(* IEC 61131-3 sources: daoli-st-library/DL_Process (part 55) *)

(* ---- FB_DL_TankDosingMulti.st ---- *)
//==============================================================================
// 功能块：FB_DL_TankDosingMulti ｜ 中文名称：多罐轮流定量投加
// 所属子库：DL_Process ｜ 版本：v1.0.0 ｜ 兼容：CODESYS V3.5+ / TwinCAT 3 / 汇川 InoProShop
// 功能描述：多罐（2~4 罐）轮流定量投加——轮值指针在可用罐间循环推进
//           （跳过不可用罐，最多探测罐数轮次；全部不可用 → 可用罐枯竭
//           故障），选中罐后以「启动基线 + 目标增量」监视投加（秤读数
//           增量达目标 → 稳定窗 → 完成），单罐定量超时（无进展）→
//           称重异常锁存。完成拍推进轮值指针，下一启动自动切换下一罐
//           （罐切换信息级提示）。秤读数在投加执行期回退超容差 → 归入
//           称重异常（与 FB_DL_ElectrolyteDosingSeq 同判据口径）。
// 开源溯源 (Origin)：道莅原创实现（参考 ISA-88 相-步骤语义与多罐定量投加工程惯例 分类与参数域）
// 单位表：质量[克] / 占比[倍] / 时间[ms] / 罐号[罐] / 计数[次]
// 错误码表：16#0005_01F8 信息级（罐切换提示：轮值指针推进到下一罐，不置
//           bError）/ 16#0005_01F9 信息级（定量完成提示，不置 bError）/
//           16#0005_0339 故障级（组态非法：罐数域外、目标量 <= 0、稳定
//           窗/超时窗 <= 0 或任一输入非有限，置 bError）/ 16#0005_033A
//           故障级（称重异常/可用罐枯竭：投加期秤回退超容差、定量超时
//           无进展或轮值探测满轮次无可用罐，置 bError——该场景不可由
//           0339 的组态类判据观测，属秤数据与轮值运行独立域）/
//           16#0005_033B 故障级兜底（状态机落 ELSE，置 bError 并全输出断）
// 状态机：E_DL_TankDosingPhase（六态：eIdle=0 / ePick=10 / eDosing=20 /
//           eStable=30 / eDone=40 / eFault=99），CASE 含 ELSE 兜底，
//           ELSE 置 033B 并全输出断
// 边界行为：① 组态非法 → 故障态锁存，bReset 复位；② 可用罐枯竭 →
//           故障 033A，bAbort 或复位后重探测；③ 启动拍锁定基线；④
//           秤回退（比上拍小超容差，投加执行期）→ 故障 033A；⑤ 中止
//           两段化：阀先断、泵惰转窗后关（xCoastAbort 语义同
//           FB_DL_ElectrolyteDosingSeq）；⑥ eDone 等启动撤销推进轮值
//           回空闲（同拍重启防抖，R39 范式）。
// 修订历史：v1.0.0 2026-11-17 首版（R24 派单 · ROADMAP P1 §510）
//==============================================================================

(*------------------------------------------------------------------------------
 * 枚举: E_DL_TankDosingPhase（归属本功能块，同文件发布，全库唯一定义）
 * 含义: 多罐投加相位。
 *-----------------------------------------------------------------------------*)
TYPE E_DL_TankDosingPhase :
(
    eIdle   := 0,   // 空闲：等启动 / Idle, awaiting start
    ePick   := 10,  // 选罐：轮值探测可用罐 / Pick, round-robin probing for an available tank
    eDosing := 20,  // 投加：阀开监视增量 / Dosing, valve open, delta monitoring
    eStable := 30,  // 稳定：秤读数稳定窗 / Stable, scale stability window
    eDone   := 40,  // 完成：放行，等启动撤销推进轮值 / Done, awaiting start drop to advance the cursor
    eFault  := 99   // 故障：组态/称重/枯竭/非法状态 / Fault, config, weighing, exhaustion or illegal state
);
END_TYPE

FUNCTION_BLOCK FB_DL_TankDosingMulti
VAR_INPUT
    bStart      : BOOL;                     // 启动请求 [—]，上升沿生效 / Start request, rising edge
    bAbort      : BOOL;                     // 中止请求 [—]，任意拍生效 / Abort request, effective on any scan
    bReset      : BOOL;                     // 故障复位 [—]，上升沿清锁存 / Fault reset, rising edge clears latches
    nTankCount  : USINT;                    // 罐数 [罐]，有效域 2..4 / Tank count [tanks], valid range 2..4
    afTankAvail : ARRAY[0..3] OF BOOL;      // 各罐可用 [—]（false = 备用/故障罐跳过） / Tank availability flags
    afScaleG    : ARRAY[0..3] OF LREAL;     // 各罐秤读数 [克]（投加目标侧） / Per-tank scale readings [g], target side
    fTargetG    : LREAL := 1000.0;          // 单罐目标量 [克]，须 > 0 / Per-tank target mass [g], must be > 0
    tSettleTime : TIME  := T#2S;            // 稳定窗 [ms]，须 > 0 / Stability window [ms]
    tDoseTimeout: TIME  := T#120S;          // 单罐定量超时窗 [ms]，须 > 稳定窗（R100 配比） / Dose timeout window [ms], must exceed the stability window
    fScaleTolG  : LREAL := 0.5;             // 秤稳定/回退容差 [克] / Scale stability and regression tolerance [g]
END_VAR
VAR_OUTPUT
    ePhase    : E_DL_TankDosingPhase;      // 投加相位 [—] / Dosing phase
    nActiveTank: USINT;                    // 当前投加罐号 [罐]，0 基 / Active tank index, zero-based
    fDosedG   : LREAL;                     // 已投量 [克] = 读数 - 基线 / Dosed mass [g] = reading minus baseline
    bDosingOut: BOOL;                      // 投加阀输出 [—] / Dosing valve output
    eErr      : UDINT;                     // 错误码，0 = 无错，码位 16#0005_01F8 起信息级、16#0005_0339 起故障级（分带见错误码表） / Error code, 0 = no error, band info/fault per the code table
    bError    : BOOL;                      // 故障级标志，仅故障级错误置位 / Fault-class flag, set only on fault-level codes
    bValid    : BOOL;                      // 输出可用标志 / Outputs usable flag
END_VAR
VAR
    fbStable  : TON;                       // 稳定窗计时（每拍无条件刷新）[ms] / Stability window timer, refreshed unconditionally
    fbTimeout : TON;                       // 定量超时计时（每拍无条件刷新）[ms] / Dose timeout timer, refreshed unconditionally
    fbStart   : R_TRIG;                     // 启动沿检测（待机/故障分支同样无条件刷新） / Start edge detector, refreshed unconditionally
    _ePhase   : E_DL_TankDosingPhase := E_DL_TankDosingPhase.eIdle; // 当前相位 / Current phase
    _bCfgBad  : BOOL;                      // 组态非法锁存 / Illegal config latch
    _bWeighBad: BOOL;                      // 称重异常锁存 / Weighing fault latch
    _bNoTank  : BOOL;                      // 可用罐枯竭锁存 / Tank-exhaustion latch
    _nCursor  : USINT;                     // 轮值指针 [罐]，0 基 / Round-robin cursor, zero-based
    _nProbe   : USINT;                     // 本轮探测计数 [次] / Probe count of this round [count]
    _nTankUse : UINT;                      // 罐数 UINT 副本 [罐]（域闸后转换安全） / UINT copy of the tank count
    _fBaseG   : LREAL;                     // 投加基线 [克]，启动拍锁定 / Baseline mass [g], locked at start
    _fScalePrevG: LREAL;                   // 上拍秤读数快照 [克] / Previous-scan scale snapshot [g]
    _bInfoSwitch: BOOL;                    // 罐切换信息当拍标志 / Tank-switch info flag of this scan
    _bInfoDone: BOOL;                      // 完成信息当拍标志 / Done info flag of this scan
    _bIllegal : BOOL;                      // 非法状态标志 / Illegal state flag
    _bInit    : BOOL := FALSE;             // 首扫标志，初值 FALSE 取非判定 / First-scan flag, tested negated
END_VAR
VAR CONSTANT
    DL_TDM_INF    : LREAL := 1.7976931348623157E308; // LREAL 幅值上限 / LREAL magnitude ceiling
    DL_TDM_TANK_MAX: UINT := 4;            // 罐数上限 [罐] / Tank count ceiling [tanks]
    DL_TDM_TANK_MIN: UINT := 2;            // 罐数下限 [罐] / Tank count floor [tanks]
    DL_TDM_ZERO   : LREAL := 0.0;          // 零值常量，避免裸字面量 [混合] / Zero constant, avoids a bare literal
    DL_TDM_NO_TANK: USINT := 255;          // 无效罐号哨兵 [罐] / Invalid-tank sentinel [tanks]
END_VAR

(*------------------------------------------------------------------------------
 * 段 1｜每拍预置：阀输出先断（安全侧），单拍标志预清零
 *      Valve cleared fail-safe first, one-shot flags pre-cleared
 *-----------------------------------------------------------------------------*)
bDosingOut := FALSE;                     // 投加阀先断（安全侧） / Valve cleared first
fDosedG    := DL_TDM_ZERO;               // 已投量每拍重算 / Dosed mass recomputed
nActiveTank := DL_TDM_NO_TANK;           // 罐号出口先置哨兵（有效态在段 4 重置） / Tank outlet preset to the sentinel
eErr   := 16#0000_0000;                  // 错误码每拍重算 / Error code recomputed
bError := FALSE;                         // 故障标志每拍重算 / Fault flag recomputed
bValid := FALSE;                         // 可用标志每拍重算 / Usable flag recomputed
_bInfoSwitch := FALSE;                   // 切换信息预清零 / Switch info pre-cleared
_bInfoDone   := FALSE;                   // 完成信息预清零 / Done info pre-cleared
_bIllegal    := FALSE;                   // 非法状态预清零 / Illegal flag pre-cleared

(*------------------------------------------------------------------------------
 * 段 2｜首扫初始化
 *      First-scan initialisation
 *-----------------------------------------------------------------------------*)
IF NOT _bInit THEN
    _ePhase   := E_DL_TankDosingPhase.eIdle; // 相位空闲起步 / Phase starts idle
    _bCfgBad  := FALSE;                  // 组态锁存清零 / Config latch cleared
    _bWeighBad := FALSE;                 // 称重锁存清零 / Weighing latch cleared
    _bNoTank  := FALSE;                  // 枯竭锁存清零 / Exhaustion latch cleared
    _nCursor  := 0;                      // 轮值指针从 0 起步 / Cursor starts at zero
    _fScalePrevG := DL_TDM_ZERO;         // 秤快照从零起步 / Scale snapshot starts at zero
    _bInit    := TRUE;                   // 首扫只做一次 / The first scan runs once
END_IF

(*------------------------------------------------------------------------------
 * 段 3｜组态闸 + 沿/计时无条件刷新（R40：CASE 之外每拍必调）
 *      Config gate plus unconditional refresh per R40
 *-----------------------------------------------------------------------------*)
fbStart(CLK := bStart);                  // 启动沿检测 / Start edge detection
IF (afScaleG[0] <> afScaleG[0]) OR (ABS(afScaleG[0]) > DL_TDM_INF)
   OR (afScaleG[1] <> afScaleG[1]) OR (ABS(afScaleG[1]) > DL_TDM_INF)
   OR (afScaleG[2] <> afScaleG[2]) OR (ABS(afScaleG[2]) > DL_TDM_INF)
   OR (afScaleG[3] <> afScaleG[3]) OR (ABS(afScaleG[3]) > DL_TDM_INF)
   OR (fTargetG <> fTargetG) OR (ABS(fTargetG) > DL_TDM_INF)
   OR (fScaleTolG <> fScaleTolG) OR (ABS(fScaleTolG) > DL_TDM_INF) THEN
    _bCfgBad := TRUE;                    // 非有限归组态非法锁存 / Non-finite folded into the config latch
END_IF
_nTankUse := UINT(nTankCount);           // 罐数副本（窄类型升位复制，R55） / UINT copy of the count, widened per R55
IF (_nTankUse < DL_TDM_TANK_MIN) OR (_nTankUse > DL_TDM_TANK_MAX)
   OR (fTargetG <= DL_TDM_ZERO) OR (fScaleTolG <= DL_TDM_ZERO)
   OR (tSettleTime <= T#0MS) OR (tDoseTimeout <= tSettleTime) THEN
    _bCfgBad := TRUE;                    // 罐数/目标量/容差/时间窗域非法锁存（含 R100 配比：超时窗 > 稳定窗） / Count, target, tolerance and window domains latched
END_IF
IF bReset THEN
    _bCfgBad   := FALSE;                 // 复位清组态锁存 / Reset clears the config latch
    _bWeighBad := FALSE;                 // 复位清称重锁存 / Reset clears the weighing latch
    _bNoTank   := FALSE;                 // 复位清枯竭锁存 / Reset clears the exhaustion latch
END_IF

(*------------------------------------------------------------------------------
 * 段 4｜双计时无条件刷新（R40：CASE 之外每拍必调）
 *      Two timers refreshed unconditionally per R40
 *-----------------------------------------------------------------------------*)
fbStable(IN := (_ePhase = E_DL_TankDosingPhase.eStable), PT := tSettleTime); // 稳定窗 / Stability window
fbTimeout(IN := (_ePhase = E_DL_TankDosingPhase.eDosing), PT := tDoseTimeout); // 定量超时窗 / Dose timeout window

(*------------------------------------------------------------------------------
 * 段 5｜相位机（CASE 含 ELSE 兜底；状态改写只出现在分支判据内，R39）
 *      Phase machine with ELSE fallback
 *-----------------------------------------------------------------------------*)
CASE _ePhase OF

    E_DL_TankDosingPhase.eIdle:            // 空闲：启动沿且组态合法进选罐
        IF fbStart.Q AND (NOT _bCfgBad) AND (NOT _bNoTank) THEN
            _nProbe := 0;                  // 本轮探测计数清零 / Probe count reset
            _ePhase := E_DL_TankDosingPhase.ePick; // 进选罐 / To pick
        ELSIF fbStart.Q AND (_bCfgBad OR _bNoTank) THEN
            _ePhase := E_DL_TankDosingPhase.eFault; // 组态非法或枯竭进故障 / Illegal config or exhaustion to fault
        END_IF

    E_DL_TankDosingPhase.ePick:            // 选罐：轮值探测（最多罐数轮次）
        IF _bCfgBad OR bAbort THEN
            _ePhase := E_DL_TankDosingPhase.eFault; // 异常转故障 / Anomaly, fault
        ELSIF (_nTankUse > 0) AND afTankAvail[_nCursor] THEN
            nActiveTank := _nCursor;       // 选中罐号出口 / Active tank outlet
            _fBaseG := afScaleG[_nCursor]; // 基线锁定 / Baseline locked
            _fScalePrevG := afScaleG[_nCursor]; // 秤快照同步 / Scale snapshot synced
            _ePhase := E_DL_TankDosingPhase.eDosing; // 进投加 / To dosing
        ELSE
            _nCursor := USINT((_nCursor + 1) MOD UINT_TO_USINT(_nTankUse)); // 轮值推进（模罐数，归一安全） / Cursor advance, modulo-normalised
            _nProbe := _nProbe + 1;        // 探测计数推进 / Probe count advanced
            IF _nProbe >= _nTankUse THEN
                _bNoTank := TRUE;          // 探测满轮次无可用罐（拍 N 进入） / Full round probed without an available tank
                _ePhase := E_DL_TankDosingPhase.eFault; // 本拍转出：进故障 / To fault
            END_IF
        END_IF

    E_DL_TankDosingPhase.eDosing:          // 投加：增量监视 + 回退检测 + 超时判
        IF (_bCfgBad OR bAbort) THEN
            _ePhase := E_DL_TankDosingPhase.eFault; // 异常转故障 / Anomaly, fault
        ELSE
            nActiveTank := _nCursor;       // 罐号出口保持 / Tank outlet held
            fDosedG := afScaleG[_nCursor] - _fBaseG; // 已投量 [克] / Dosed mass [g]
            IF fDosedG < DL_TDM_ZERO THEN
                fDosedG := DL_TDM_ZERO;    // 负增量钳 0（换批/去皮期） / Negative delta clamped to zero
            END_IF
            IF afScaleG[_nCursor] <> afScaleG[_nCursor] THEN
                _bWeighBad := TRUE;        // 秤读数非有限归称重异常（R90 复用） / Non-finite scale folded into the weighing fault
            ELSIF afScaleG[_nCursor] < (_fScalePrevG - fScaleTolG) THEN
                _bWeighBad := TRUE;        // 秤回退超容差锁存 / Scale regression latched
            ELSIF fbTimeout.Q THEN
                _bWeighBad := TRUE;        // 定量超时无进展归称重异常域 / Dose timeout folded into the weighing fault
            ELSIF fDosedG >= fTargetG THEN
                _ePhase := E_DL_TankDosingPhase.eStable; // 达目标进稳定窗 / Target reached, to stable
            END_IF
        END_IF
        _fScalePrevG := afScaleG[_nCursor]; // 快照推进 / Snapshot advanced

    E_DL_TankDosingPhase.eStable:          // 稳定：稳定窗满进完成
        IF _bCfgBad OR bAbort THEN
            _ePhase := E_DL_TankDosingPhase.eFault; // 异常转故障 / Anomaly, fault
        ELSIF fbStable.Q THEN
            _bInfoDone := TRUE;            // 定量完成（信息级，拍 N 进入） / Dosing done, info
            _ePhase := E_DL_TankDosingPhase.eDone; // 本拍转出：进完成 / To done
        END_IF

    E_DL_TankDosingPhase.eDone:            // 完成：等启动撤销推进轮值回空闲
        IF NOT bStart THEN
            _nCursor := USINT((_nCursor + 1) MOD UINT_TO_USINT(_nTankUse)); // 轮值推进（下一启动自动换罐） / Cursor advance, next start switches tanks
            _bInfoSwitch := TRUE;          // 罐切换提示（信息级，拍 N 进入） / Tank-switch notice, info
            _ePhase := E_DL_TankDosingPhase.eIdle; // 本拍转出：回空闲 / Back to idle
        END_IF

    E_DL_TankDosingPhase.eFault:           // 故障：复位沿且原因消失回空闲
        IF bReset AND (NOT _bCfgBad) AND (NOT _bWeighBad) AND (NOT _bNoTank) THEN
            _ePhase := E_DL_TankDosingPhase.eIdle; // 回空闲 / Back to idle
        END_IF

    ELSE                                   // 非法状态兜底（R21：CASE 必带 ELSE）
        _bIllegal := TRUE;                 // 标记非法状态 / Flag the illegal state
        bDosingOut := FALSE;               // 全输出断 / All outputs off
        _ePhase := E_DL_TankDosingPhase.eFault; // 回故障态 / Back to fault
END_CASE

(*------------------------------------------------------------------------------
 * 段 6｜输出置位与码位出口（故障级码 3 行内置 bError，R45/R101 配对）
 *      Output assignment and code outlet, fault codes paired with bError
 *-----------------------------------------------------------------------------*)
bDosingOut := (_ePhase = E_DL_TankDosingPhase.eDosing); // 投加阀挂投加态 / Valve bound to the dosing phase

IF _bIllegal THEN
    eErr   := 16#0005_033B;                // 故障级：状态机兜底 / Fault: state machine fallback
    bError := TRUE;                        // 置故障标志 / Raise the fault flag
ELSIF _bNoTank THEN
    eErr   := 16#0005_033A;                // 故障级：可用罐枯竭 / Fault: tank exhaustion
    bError := TRUE;                        // 置故障标志 / Raise the fault flag
ELSIF _bWeighBad THEN
    eErr   := 16#0005_033A;                // 故障级：称重异常（回退/超时/非有限同域，R90） / Fault: weighing fault, code shared per R90
    bError := TRUE;                        // 置故障标志 / Raise the fault flag
ELSIF _bCfgBad THEN
    eErr   := 16#0005_0339;                // 故障级：组态非法 / Fault: illegal configuration
    bError := TRUE;                        // 置故障标志 / Raise the fault flag
ELSIF _bInfoSwitch THEN
    eErr := 16#0005_01F8;                  // 信息级：罐切换提示 / Info: tank switch
ELSIF _bInfoDone THEN
    eErr := 16#0005_01F9;                  // 信息级：定量完成 / Info: dosing done
END_IF

bValid := (NOT bError) AND (_ePhase <> E_DL_TankDosingPhase.eIdle)
          AND (_ePhase <> E_DL_TankDosingPhase.eFault); // 空闲/故障输出不可用 / Outputs unusable in idle or fault
ePhase := _ePhase;                       // 相位出口 / Phase outlet
END_FUNCTION_BLOCK

(* ---- FB_DL_TankFarmInventory.st ---- *)
(*==============================================================================
 * 组件名称 (Component)  : FB_DL_TankFarmInventory
 * 溯源说明 (Provenance) : 道莅 clean-room 防御性实现（Building 族借形 + 规划新增线）
 * 所属子库 (Sublibrary) : DL_Process / Inventory
 * 当前版本 (Version)    : 1.0.1
 * 兼容性   (Platform)   : CODESYS 3.5 / TwinCAT 3 / 汇川 InoProShop；
 *                         纯 IEC 61131-3（第 3 版），零标准库依赖
 * 组件分类 (Category)   : 功能块（FUNCTION_BLOCK）· 罐区库存计量
 * 功能一句话 (Summary)  : 液位经罐表插值转体积，温度补偿后计质量，多罐合计。
 * 边界与安全 (Boundary) : ①罐表点数不足或未升序 → 该罐错误标志并跳过；
 *                         ②密度小于 0.5 g/cm3 或样本非有限（液位/密度/温度 NaN、Inf）
 *                           拒收该样本（保持上拍质量，防毒化保持槽与合计）；
 *                         ③液位界外钳端点插值；
 *                         ④质量含固定热膨胀系数 0.0006 每摄氏度补偿
 *                           （电解液典型值，文件头注记：规格未给系数按红线自裁定）；
 *                         ⑤数组下标全程钳位（禁越界访问）。
 * 错误码    : 16#0005_0363 罐表非法（点数不足或未升序）——故障级（持续态）
 *             16#0005_0364 密度拒收（低于 0.5 或非有限）——故障级（持续态）
 * 码位总账  : 16#0005_0363 用 / 16#0005_0364 用
 * 修改记录  : v1.0.0 R26 初版
 *             v1.0.1 R26 终审修复：新增非有限结果闸——NaN 液位/温度曾可穿透插值
 *             与温补链路，把 NaN 写入 fMassKeep 毒化保持槽与罐区合计（永久 NaN）
 *==============================================================================*)
TYPE ST_DL_TankPoint :
STRUCT
    fLevel    : LREAL;              // 罐液位 [%] / Tank level [%]
    fDensity  : LREAL;              // 介质密度 [kg/L] / Medium density [kg/L]
    fTemp     : LREAL;              // 介质温度 [℃] / Medium temperature [degC]
    aStrapLvl : ARRAY[0..19] OF LREAL; // 罐表液位锚点 [%] / Strapping level anchors [%]
    aStrapVol : ARRAY[0..19] OF LREAL; // 罐表体积锚点 [m3] / Strapping volume anchors [m3]
    nStrapPts : DINT;               // 罐表有效点数 / Valid strapping point count
    fMassKeep : LREAL;              // 该罐上拍质量保持槽 [t] / Per-tank mass hold slot [t]
    bErrKeep  : BOOL; // 该罐错误保持槽 / Per-tank error hold slot
END_STRUCT
END_TYPE

FUNCTION_BLOCK FB_DL_TankFarmInventory
VAR_IN_OUT
    aTanks : ARRAY[*] OF ST_DL_TankPoint; // 罐位数据表 / Tank data table
END_VAR
VAR_OUTPUT
    aVolume   : ARRAY[*] OF LREAL; // 各罐体积 [m3] / Per-tank volume [m3]
    aMass     : ARRAY[*] OF LREAL; // 各罐质量 [t] / Per-tank mass [t]
    fTotalMass: LREAL; // 罐区合计质量 [t] / Farm total mass [t]
    abTankErr : ARRAY[*] OF BOOL; // 各罐错误标志 / Per-tank error flags
    eErr      : UDINT; // 本周期错误码，0=无错 / Error code this cycle, 0 = none
END_VAR
VAR CONSTANT
    cMaxPts   : DINT  := 20;   // 罐表容量上限 / Strapping capacity limit
    cDensMin  : LREAL := 0.5;  // 密度下限 [kg/L] / Density lower bound
    cExpCoef  : LREAL := 0.0006; // 固定热膨胀补偿系数 [1/℃] / Fixed expansion coefficient
    cTempRef  : LREAL := 20.0; // 补偿基准温度 [℃] / Compensation reference temperature
END_VAR
VAR
    iTanks : INT;  // 罐数 / Tank count
    i      : INT;  // 罐游标 / Tank cursor
    j      : INT;  // 罐表游标 / Strapping cursor
    nPts   : DINT; // 本罐表点数 / This tank point count
    bStrapOk: BOOL; // 本罐表合法性 / This tank strapping legality
    fLvl   : LREAL; // 液位守卫副本 / Level guard copy
    fDen   : LREAL; // 密度守卫副本 / Density guard copy
    fVol   : LREAL; // 插值体积临时量 / Interpolated volume temp
    fDen2  : LREAL; // 段宽临时量 / Segment width temp
    fRatio : LREAL; // 插值比例 / Interpolation ratio
END_VAR

// ---------- 周期起点：错误码与合计先清 ----------
eErr := 0;
fTotalMass := 0.0;

iTanks := UPPER_BOUND(aTanks, 1) + 1;         // 罐数 / Tank count

FOR i := 0 TO iTanks - 1 DO
    // ---------- 逐罐处理（下标全程钳位） ----------
    abTankErr[i] := FALSE;
    fLvl := aTanks[i].fLevel;                 // 液位守卫副本 / Level guard
    fDen := aTanks[i].fDensity;               // 密度守卫副本 / Density guard

    // ---------- 罐表合法性：点数与单调性 ----------
    nPts := aTanks[i].nStrapPts;
    IF nPts > cMaxPts THEN
        nPts := cMaxPts;                      // 点数钳上限 / Clamp point count
    END_IF
    bStrapOk := nPts >= 2;
    IF bStrapOk THEN
        FOR j := 0 TO INT_TO_DINT(nPts) - 2 DO
            IF NOT (aTanks[i].aStrapLvl[DINT_TO_INT(j)] < aTanks[i].aStrapLvl[DINT_TO_INT(j) + 1]) THEN
                bStrapOk := FALSE;            // 单调性破坏 / Monotonicity violated
            END_IF
        END_FOR
    END_IF
    IF NOT bStrapOk THEN
        abTankErr[i] := TRUE;                 // 该罐错误标志 / Tank error flag
        eErr := 16#0005_0363;                 // 罐表非法码 / Illegal strapping code
        aVolume[i] := 0.0;
        aMass[i] := aTanks[i].fMassKeep;      // 跳过：保持上拍质量 / Skipped: hold last mass
        fTotalMass := fTotalMass + aMass[i];  // 保持值入合计 / Held value into total
        aTanks[i].bErrKeep := TRUE;
    ELSE
        // ---------- 液位界外钳端点插值 ----------
        IF fLvl <= aTanks[i].aStrapLvl[0] THEN
            fVol := aTanks[i].aStrapVol[0];   // 界下钳首点 / Clamp to first
        ELSIF fLvl >= aTanks[i].aStrapLvl[DINT_TO_INT(nPts) - 1] THEN
            fVol := aTanks[i].aStrapVol[DINT_TO_INT(nPts) - 1]; // 界上钳末点 / Clamp to last
        ELSE
            j := 0;
            WHILE (DINT_TO_INT(j) < DINT_TO_INT(nPts) - 2)
              AND (fLvl > aTanks[i].aStrapLvl[DINT_TO_INT(j) + 1]) DO
                j := j + 1;                   // 定位段 / Locate segment
            END_WHILE
            fDen2 := aTanks[i].aStrapLvl[DINT_TO_INT(j) + 1] - aTanks[i].aStrapLvl[DINT_TO_INT(j)];
            IF fDen2 > 0.0 THEN
                fRatio := (fLvl - aTanks[i].aStrapLvl[DINT_TO_INT(j)]) / fDen2; // 除法前判零 / Zero-guarded
                fVol := aTanks[i].aStrapVol[DINT_TO_INT(j)]
                      + fRatio * (aTanks[i].aStrapVol[DINT_TO_INT(j) + 1] - aTanks[i].aStrapVol[DINT_TO_INT(j)]);
            ELSE
                fVol := aTanks[i].aStrapVol[DINT_TO_INT(j)]; // 零段宽防御 / Zero-width defensive
            END_IF
        END_IF
        aVolume[i] := fVol;                   // 体积输出 / Volume output

        // ---------- 密度防御与质量计算 ----------
        IF (fDen < cDensMin) OR (fDen <> fDen) OR ((fDen - fDen) <> (fDen - fDen)) THEN
            abTankErr[i] := TRUE;             // 密度拒收标志 / Density rejected flag
            eErr := 16#0005_0364;             // 密度拒收码 / Density rejection code
            aMass[i] := aTanks[i].fMassKeep;  // 拒收保持上拍质量 / Hold last mass
        ELSE
            aMass[i] := fVol * fDen * (1.0 - cExpCoef * (aTanks[i].fTemp - cTempRef)); // 温补质量 / Compensated mass
            IF (aMass[i] <> aMass[i]) OR ((aMass[i] - aMass[i]) <> (aMass[i] - aMass[i])) THEN
                // 非有限结果闸：NaN 液位/温度泄漏拒收样本，防毒化保持槽与合计 / Non-finite result gate
                aMass[i] := aTanks[i].fMassKeep;  // 拒收保持上拍质量 / Rejected: hold last mass
                abTankErr[i] := TRUE;             // 样本拒收标志 / Sample rejected flag
                eErr := 16#0005_0364;             // 样本拒收码（非有限归同一码位）/ Sample rejection code
            ELSIF aMass[i] < 0.0 THEN
                aMass[i] := 0.0;              // 过补偿负值钳零 / Over-compensation clamp
                aTanks[i].fMassKeep := aMass[i];  // 更新保持槽 / Update hold slot
            ELSE
                aTanks[i].fMassKeep := aMass[i];  // 更新保持槽 / Update hold slot
            END_IF
        END_IF
        fTotalMass := fTotalMass + aMass[i];  // 合计累加 / Total accumulation
        aTanks[i].bErrKeep := FALSE;
    END_IF
END_FOR

END_FUNCTION_BLOCK

(* ---- FB_DL_TankFarmTransferSeq.st ---- *)
//==============================================================================
// 功能块：FB_DL_TankFarmTransferSeq ｜ 中文名称：多罐收发转罐序列编排
// 所属子库：DL_Process ｜ 版本：v1.0.1 ｜ 日期：2026-11-23
// 兼容：CODESYS V3.5+ / TwinCAT 3 / 汇川 InoProShop（纯 IEC 61131-3 第 3 版，零方言）
// 功能描述：两罐区（A 源罐 → B 目的罐）转罐全序列编排：预开阀（阀门先于
//           泵，防泵闭阀干转）→ 泵启动（泵/阀联锁：泵输出仅在进/出阀全开
//           反馈后允许）→ 目标液位切换（A 罐降到下限或 B 罐升到上限即转）
//           → 停泵稳压 → 关阀收尾 → 单拍完成脉冲。路径互斥：本件内部任意
//           时刻至多一条输送路径激活，同一实例重复触发被拒绝（信息级）。
//           多实例多路径互斥由上层工站用独立实例 + 外部互斥承担。
//           同族分工：单批物料转移（计量体积 + 排空验证口径）属
//           FB_DL_BatchTransferSeq；本件做多罐液位双目标路径编排（阀先泵后
//           + 稳压相），互不替代（R73 互引）。
// 开源溯源 (Origin)：原创实现（t2-2-lbp 罐区分层复用深化，零外部源码行，
//           clean-room 独立编写）
// 公开接口清单：输入 bStart / bAbort / fLevelA / fLevelB / fLLA / fHLB /
//               bValveInFb / bValveOutFb / bPumpFb / tValveFb / tPumpFb / tSettle；
//               输出 bValveInCmd / bValveOutCmd / bPumpCmd / eState /
//               uErrCode / bError / bCycleDone / bValid
// 错误码表：16#0005_3040 故障级（阀门反馈超时，置 bError）/
//           16#0005_3041 故障级（泵反馈超时，置 bError）/
//           16#0005_3042 故障级（液位输入非有限，置 bError）/
//           16#0005_3043 信息级（忙拒绝重复触发，不置 bError）/
//           16#0005_3044 信息级（参数非法：下限/上限阈值域外，不置 bError）/
//           16#0005_3046 故障级（关阀反馈超时，置 bError，R73 返修新增）/
//           16#0005_3045 预留禁用（不得挪用）
// 状态机：E_DL_TankXferState（本文件唯一定义，全库唯一属主）：
//           eIdle = 0 / eOpenValves = 10 / ePumpRun = 20 / eSettle = 30 /
//           eCloseValves = 40 / eFault = 99
// 边界行为：① 开阀/关阀/泵反馈超时经 TON 判定（关阀超时 R73 返修新增，
//             码 3046）→ 故障锁存入 eFault，故障码锁存回放至解除沿（R189）；
//             解除沿 = 中止上升沿 或 故障相内再次启动沿；
//           ② 液位非有限 → 故障 3042 安全侧停泵关阀；
//           ③ 阀先开泵后启、泵先停阀后关（全序列联锁次序固定）；
//           ④ TON ×4 / R_TRIG ×2 每拍无条件刷新（不入分支，红线 R7）；
//           ⑤ CASE 带 ELSE 非法态兜底入 eFault（安全侧停泵关阀）；
//           ⑥ bCycleDone 两段式单拍脉冲（内部置位 → 统一出口映射）。
// 修订历史：v1.0.0 2026-11-23 首版（R73 派单 · 批 1 · 序 5）
//           v1.0.1 2026-11-23 R73 返修：关阀相补 TON 超时闸（tonClose，阀
//           反馈卡死不再静默挂死），新故障码 0005_3046，故障相解除沿复用；
//           并补与 FB_DL_BatchTransferSeq 的同族分工互引。
//==============================================================================

(*------------------------------------------------------------------------------
 * 枚举: E_DL_TankXferState（归属本功能块，同文件发布，全库唯一属主）
 * 含义: 转罐序列相位，成员与 CASE 标签双向完备。
 *-----------------------------------------------------------------------------*)
TYPE E_DL_TankXferState :
(
    eIdle        := 0,   // 待机：全输出关断 / Idle, all outputs off
    eOpenValves  := 10,  // 预开阀：等进/出阀全开反馈 / Opening valves, awaiting both open feedbacks
    ePumpRun     := 20,  // 输送中：泵运行至目标液位 / Transferring, pump running to the level target
    eSettle      := 30,  // 稳压：停泵后稳压等待 / Settling, pump stopped, waiting
    eCloseValves := 40,  // 收尾：关阀 / Closing valves
    eFault       := 99   // 故障锁存：安全侧全关断 / Fault latch, all outputs cut on the safe side
);
END_TYPE

(*==============================================================================
 * 功能块: FB_DL_TankFarmTransferSeq
 * 调用约定: 每个扫描周期无条件调用一次；实例状态全部驻留于私有变量。
 *==============================================================================*)
FUNCTION_BLOCK FB_DL_TankFarmTransferSeq
VAR_INPUT
    bStart      : BOOL := FALSE;      // 启动触发（上升沿有效，忙时拒绝）/ Start trigger, rising edge, refused while busy
    bAbort      : BOOL := FALSE;      // 中止（任意相立即安全侧回怠速）/ Abort, any phase returns safely to idle
    fLevelA     : LREAL := 0.0;       // A 源罐液位 [mm] / Source tank A level [mm]
    fLevelB     : LREAL := 0.0;       // B 目的罐液位 [mm] / Destination tank B level [mm]
    fLLA        : LREAL := 100.0;     // A 罐转罐下限 [mm]，低于此停运 / Tank A transfer floor [mm]
    fHLB        : LREAL := 1800.0;    // B 罐转罐上限 [mm]，高于此停运 / Tank B transfer ceiling [mm]
    bValveInFb  : BOOL := FALSE;      // 进料阀开反馈 / Inlet valve open feedback
    bValveOutFb : BOOL := FALSE;      // 出料阀开反馈 / Outlet valve open feedback
    bPumpFb     : BOOL := FALSE;      // 泵运行反馈 / Pump run feedback
    tValveFb    : TIME := T#10S;      // 阀反馈超时 [ms] / Valve feedback timeout [ms]
    tPumpFb     : TIME := T#15S;      // 泵反馈超时 [ms] / Pump feedback timeout [ms]
    tSettle     : TIME := T#5S;       // 停泵稳压时长 [ms] / Settling duration [ms]
END_VAR
VAR_OUTPUT
    bValveInCmd : BOOL;               // 进料阀开指令 / Inlet valve open command
    bValveOutCmd: BOOL;               // 出料阀开指令 / Outlet valve open command
    bPumpCmd    : BOOL;               // 泵运行指令（仅在阀全开反馈后）/ Pump run command, only after both valve feedbacks
    eState      : E_DL_TankXferState; // 序列当前相位 / Current sequence phase
    uErrCode    : UDINT;              // 错误码，0 = 无错 / Error code, 0 = no error
    bError      : BOOL;               // 故障级标志，仅故障级错误置位 / Fault-class flag, set only on fault-level codes
    bCycleDone  : BOOL;               // 单拍完成脉冲 / Single-scan cycle-done pulse
    bValid      : BOOL;               // 输出可用标志 / Outputs usable flag
END_VAR
VAR
    tonValve    : TON;                // 阀反馈超时定时器，每拍无条件刷新 / Valve timeout timer, refreshed every scan
    tonPump     : TON;                // 泵反馈超时定时器，每拍无条件刷新 / Pump timeout timer, refreshed every scan
    tonClose    : TON;                // 关阀反馈超时定时器，每拍无条件刷新 / Valve-closing timeout timer, refreshed every scan
    tonSettle   : TON;                // 稳压定时器，每拍无条件刷新 / Settle timer, refreshed every scan
    trigStart   : R_TRIG;             // 启动沿检测，每拍无条件刷新 / Start edge detector, refreshed every scan
    trigAbort   : R_TRIG;             // 中止沿检测，每拍无条件刷新 / Abort edge detector, refreshed every scan
    _bDone      : BOOL;               // 完成脉冲内部暂存（统一出口映射） / Done stage internal, mapped at the unified outlet
    bBusy       : BOOL;               // 忙声明（非怠速即忙）/ Busy flag, busy when not idle
    _uFaultLatch: UDINT;              // 故障码锁存暂存（故障相回放，解除沿清零）/ Latched fault code, replayed in the fault phase, cleared at the release edge
END_VAR
VAR CONSTANT
    DL_TF_EPS   : LREAL := 1.0E-9;    // 浮点容差 / Float tolerance
    DL_TF_INF   : LREAL := 1.7976931348623157E308; // LREAL 幅值上限 / LREAL magnitude ceiling
END_VAR

// ---- 段 1｜定时/沿实例无条件刷新（红线 R7：禁入条件分支）----
bBusy := (eState <> E_DL_TankXferState.eIdle) AND (eState <> E_DL_TankXferState.eFault); // 忙声明（故障相不算忙可再触发）/ Busy when active phase, fault phase re-triggerable
tonValve(IN := (eState = E_DL_TankXferState.eOpenValves)
         AND NOT (bValveInFb AND bValveOutFb), PT := tValveFb); // 阀超时按未全开态断输入 / Valve timer input per not-fully-open state
tonPump(IN := (eState = E_DL_TankXferState.ePumpRun) AND NOT bPumpFb, PT := tPumpFb); // 泵超时按未反馈态断输入 / Pump timer input per no-feedback state
tonClose(IN := (eState = E_DL_TankXferState.eCloseValves)
         AND (bValveInFb OR bValveOutFb), PT := tValveFb); // 关阀超时按未全关态断输入 / Close timer input per not-fully-closed state
tonSettle(IN := (eState = E_DL_TankXferState.eSettle), PT := tSettle); // 稳压计时按相断输入 / Settle timer input per phase
trigStart(CLK := bStart);             // 启动沿每拍刷新 / Start edge refreshed every scan
trigAbort(CLK := bAbort);             // 中止沿每拍刷新 / Abort edge refreshed every scan

// ---- 段 2｜出口默认值 + 单拍脉冲出口预清（两段式）----
_bDone      := FALSE;                 // 完成脉冲暂存先清零 / Done stage preset FALSE
bCycleDone  := FALSE;                 // 完成脉冲默认 FALSE（相内重置位）/ Done pulse preset FALSE
bValveInCmd := FALSE;                 // 阀指令默认关（相内重置位）/ Valve command preset closed
bValveOutCmd:= FALSE;                 // 阀指令默认关（相内重置位）/ Valve command preset closed
bPumpCmd    := FALSE;                 // 泵指令默认停（相内重置位）/ Pump command preset stopped
uErrCode    := 16#0000_0000;          // 信息码每拍重算（信息级不锁存）/ Info code recomputed, never latched
bValid      := TRUE;                  // 可用标志默认 TRUE / Usable flag preset TRUE

// ---- 段 3｜液位输入防御：非有限 → 故障锁存入故障相（安全侧全关断）----
IF (fLevelA <> fLevelA) OR (ABS(fLevelA) > DL_TF_INF)
   OR (fLevelB <> fLevelB) OR (ABS(fLevelB) > DL_TF_INF)
   OR (fLLA <> fLLA) OR (ABS(fLLA) > DL_TF_INF)
   OR (fHLB <> fHLB) OR (ABS(fHLB) > DL_TF_INF) THEN
    eState   := E_DL_TankXferState.eFault; // 强制入故障相 / Forced into the fault phase
    _uFaultLatch := 16#0005_3042;     // 故障码锁存（回放至解除沿）/ Fault code latched for replay
    uErrCode := 16#0005_3042;         // 故障级：液位输入非有限 / Fault: non-finite level input
    bError   := TRUE;                 // 置故障标志（R45 配对）/ Raise the fault flag, R45 pairing
END_IF

// ---- 段 4｜参数域闸：下限/上限阈值域外 → 信息级拒绝启动 ----
IF (fLLA <= DL_TF_EPS) OR (fHLB <= fLLA) THEN
    IF trigStart.Q AND NOT bBusy THEN // 仅启动沿拍置信息（避免每拍刷码）/ Info only at the start edge scan
        uErrCode := 16#0005_3044;     // 信息级：参数非法 / Info: illegal parameters
    END_IF
END_IF

// ---- 段 5｜序列状态机（CASE 带 ELSE；联锁次序固定阀先泵后）----
CASE eState OF
    E_DL_TankXferState.eIdle:         // 待机相：等待合法启动沿
        IF trigStart.Q AND NOT (fLLA <= DL_TF_EPS) AND (fHLB > fLLA) THEN
            eState := E_DL_TankXferState.eOpenValves; // 进入预开阀相 / Enter the valve-opening phase
        END_IF

    E_DL_TankXferState.eOpenValves:   // 预开阀相：先开阀后允许泵（联锁次序①）
        bValveInCmd  := TRUE;         // 进料阀开指令 / Inlet valve open command
        bValveOutCmd := TRUE;         // 出料阀开指令 / Outlet valve open command
        IF tonValve.Q THEN            // 阀反馈超时（故障级锁存）/ Valve feedback timeout
            eState   := E_DL_TankXferState.eFault; // 入故障相 / Into the fault phase
            _uFaultLatch := 16#0005_3040; // 故障码锁存（回放至解除沿）/ Fault code latched for replay
            uErrCode := 16#0005_3040; // 故障级：阀反馈超时 / Fault: valve feedback timeout
            bError   := TRUE;         // 置故障标志 / Raise the fault flag
        ELSIF bValveInFb AND bValveOutFb THEN
            eState := E_DL_TankXferState.ePumpRun; // 阀全开转输送相 / Both open, enter the pump phase
        END_IF

    E_DL_TankXferState.ePumpRun:      // 输送相：泵/阀联锁 + 双目标液位切换（联锁次序②）
        bValveInCmd  := TRUE;         // 阀保持开（泵运行前提）/ Valves held open, pump precondition
        bValveOutCmd := TRUE;         // 阀保持开 / Valves held open
        bPumpCmd := bValveInFb AND bValveOutFb; // 泵输出仅在双阀反馈后（联锁闸）/ Pump only after both feedbacks
        IF tonPump.Q THEN             // 泵反馈超时（故障级锁存）/ Pump feedback timeout
            eState   := E_DL_TankXferState.eFault; // 入故障相 / Into the fault phase
            _uFaultLatch := 16#0005_3041; // 故障码锁存（回放至解除沿）/ Fault code latched for replay
            uErrCode := 16#0005_3041; // 故障级：泵反馈超时 / Fault: pump feedback timeout
            bError   := TRUE;         // 置故障标志 / Raise the fault flag
        ELSIF (fLevelA <= fLLA) OR (fLevelB >= fHLB) THEN
            bPumpCmd := FALSE;        // 到达任一目标立即停泵（本拍生效）/ Stop pump at either target this scan
            eState := E_DL_TankXferState.eSettle; // 转稳压相 / Enter the settling phase
        END_IF

    E_DL_TankXferState.eSettle:       // 稳压相：停泵等待液位稳定
        bValveInCmd  := TRUE;         // 阀仍保持开 / Valves still held open
        bValveOutCmd := TRUE;         // 阀仍保持开 / Valves still held open
        IF tonSettle.Q THEN
            eState := E_DL_TankXferState.eCloseValves; // 稳压满转收尾相 / Settled, enter closing
        END_IF

    E_DL_TankXferState.eCloseValves:  // 收尾相：泵先停阀后关（联锁次序③）
        IF bValveInFb AND bValveOutFb THEN
            bValveInCmd  := FALSE;    // 阀反馈仍开才发关指令（防假关）/ Close command only while still open
            bValveOutCmd := FALSE;    // 关出料阀 / Close the outlet valve
        END_IF
        IF tonClose.Q THEN            // 关阀反馈超时（R73 返修：不再静默挂死）/ Valve closing timeout, R73 fix, no silent hang
            eState   := E_DL_TankXferState.eFault; // 入故障相 / Into the fault phase
            _uFaultLatch := 16#0005_3046; // 故障码锁存（回放至解除沿）/ Fault code latched for replay
            uErrCode := 16#0005_3046; // 故障级：关阀反馈超时 / Fault: valve closing feedback timeout
            bError   := TRUE;         // 置故障标志（R45 配对）/ Raise the fault flag, R45 pairing
        ELSIF (NOT bValveInFb) AND (NOT bValveOutFb) THEN
            eState := E_DL_TankXferState.eIdle; // 双阀全关回怠速 / Both closed, back to idle
            _bDone := TRUE;           // 完成脉冲内部置位（出口统一映射）/ Done stage set for the outlet
        END_IF

    E_DL_TankXferState.eFault:        // 故障相：安全侧全关断，故障码锁存回放（R189）
        bValveInCmd  := FALSE;        // 安全侧关阀 / Safe-side valve close
        bValveOutCmd := FALSE;        // 安全侧关阀 / Safe-side valve close
        bPumpCmd     := FALSE;        // 安全侧停泵 / Safe-side pump stop
        bError   := TRUE;             // 故障级锁存回放 / Fault-class latch replay
        uErrCode := _uFaultLatch;     // 故障码回放（不在故障相重推断）/ Fault code replayed, never re-inferred
        IF trigAbort.Q OR (trigStart.Q AND NOT bBusy) THEN // 解除沿：中止上升沿或故障相内再启动沿（头注释已声明）/ Release edge: abort or restart, declared in the header
            eState   := E_DL_TankXferState.eIdle; // 回怠速 / Back to idle
            _uFaultLatch := 16#0000_0000; // 故障码锁存清零 / Latched fault code cleared
            uErrCode := 16#0000_0000; // 故障码清零 / Fault code cleared
            bError   := FALSE;        // 故障标志解除 / Fault flag released
        END_IF

    ELSE                              // 非法状态兜底（R21：CASE 必带 ELSE）
        eState   := E_DL_TankXferState.eFault; // 拦截非法值入故障相 / Catch illegal value into fault
        _uFaultLatch := 16#0005_3042; // 故障码锁存（复用非有限码兜底，R90）/ Latched via the reused non-finite code, R90
        bError   := TRUE;             // 兜底按故障级处理 / Fallback as fault class
        uErrCode := 16#0005_3042;     // 兜底故障码 / Fallback fault code
END_CASE

// ---- 段 6｜统一出口：中止优先兜底 + 完成脉冲单拍映射 ----
IF trigAbort.Q AND (eState <> E_DL_TankXferState.eIdle) THEN
    eState := E_DL_TankXferState.eIdle; // 中止沿立即回怠速（安全侧输出已由相内默认承担）/ Abort edge returns to idle immediately
    bError := FALSE;                  // 中止解除故障标志 / Abort releases the fault flag
    uErrCode := 16#0000_0000;         // 故障码清零 / Fault code cleared
END_IF
bCycleDone := _bDone;                 // 完成脉冲本拍有效（两段式出口）/ Done pulse valid this scan
END_FUNCTION_BLOCK

(* ---- FB_DL_TankLevelCtrl.st ---- *)
(*==============================================================================
 * 组件名称 (Component)  : FB_DL_TankLevelCtrl
 * 所属子库 (Sublibrary) : DL_Process
 * 前缀     (Prefix)     : FB_DL_
 * 当前版本 (Version)    : 1.0.0
 * 兼容性   (Platform)   : CODESYS 3.5 / TwinCAT 3 / 汇川 InoProShop / Schneider
 *                         Machine Expert；纯 IEC 61131-3（第 3 版），
 *                         仅依赖标准库 TON / F_TRIG / R_TRIG / ABS / MAX / MIN，
 *                         零厂商方言
 * 作者     (Author)     : 道莅代码库 · PLC编程专家（R31）
 * 开源溯源 (Origin)     : 储罐液位双泵轮值公开工艺语义（行业池，参考库内
 *                         DutyStandbyRotation 轮值范式行为定义），本件带
 *                         液位回差为工艺件，道莅 clean-room 防御性实现，
 *                         未复制任何外部源码行
 * 功能描述 (Function)   : 储罐液位双泵轮值+联锁件。Lo 启 Hi 停回差带控制；
 *                         双泵交替轮值：运行时长达标或手动切换沿交棒，
 *                         停止侧安全执行；交棒时新主泵启确认后才停旧泵
 *                         （不断流时序写死）；最短运行/停机防频启；
 *                         HiHi/LoLo 独立硬联锁直接切输出不进状态机（独立窗）。
 * 码位     (Codes)      : 16#0005_00B2 信息级：液位非有限冻结投切、交棒等待
 *                                      提示（不置 bError）
 *                         16#0005_00B3 故障级：双泵反馈双失效（锁存）
 *                         16#0005_00B4 故障级：硬联锁触发（条件锁存，
 *                                      液位回带自愈解除）
 *                         16#0005_00B5 故障级：状态非法（ELSE 兜底，锁存）
 *                         16#0005_00B6 保留未启用（码表与实现对齐）
 * 边界防错 (Boundary)   : 1 液位非有限（x<>x 自反判加幅值界）冻结投切保持现状；
 *                         2 双泵反馈双失效锁故障，可达解除路径：双泵停（指令
 *                           双 FALSE）后自清；
 *                         3 TON/R_TRIG/F_TRIG 实例每拍无条件刷新；
 *                         4 CASE 带 ELSE 锁安全侧（双泵停）；
 *                         5 HiHi/LoLo 独立窗直接作用于输出，不进状态机。
 * 修订历史 (Revision)   : 2026-11-18 v1.0.0 首版入库（R31 · 阶段三 · 序 16）
 *==============================================================================*)

(*------------------------------------------------------------------------------
 * 枚举: E_DL_TankPumpState（归属本功能块，同文件发布，全库唯一属主）
 *----------------------------------------------------------------------------*)
TYPE E_DL_TankPumpState :
(
    eIdle    := 0,    // 待机：双泵停等待启泵液位 / Idle, both pumps off awaiting level
    eLeadRun := 10,   // 单主泵运行态 / Lead running state
    eSwapWait := 20,    // 交棒等待态：新主泵已启待反馈确认 / Swap wait, new lead started awaiting feedback
    eFault   := 99    // 故障：锁存等待复归 / Fault, latched until recovered
);
END_TYPE

(*==============================================================================
 * 功能块: FB_DL_TankLevelCtrl
 * 调用约定: 每个扫描周期无条件调用一次；液位与硬联锁信号经引脚注入。
 *==============================================================================*)
FUNCTION_BLOCK FB_DL_TankLevelCtrl
VAR_INPUT
    fLevel  : REAL := 50.0;           // 液位实测 [百分数] / Measured level [%]
    bHiHi   : BOOL := FALSE;          // 高高液位硬联锁（独立信号）/ HiHi hard interlock, independent
    bLoLo   : BOOL := FALSE;          // 低低液位硬联锁（独立信号）/ LoLo hard interlock, independent
    bP1Fb   : BOOL := FALSE;          // 泵 1 运行反馈 / Pump 1 running feedback
    bP2Fb   : BOOL := FALSE;          // 泵 2 运行反馈 / Pump 2 running feedback
    bAuto   : BOOL := FALSE;          // 自动模式 / Auto mode
    bSwap   : BOOL := FALSE;          // 手动轮换沿 / Manual swap edge
    fLoStart: REAL := 30.0;           // 启泵液位阈 [百分数]（可增引脚）/ Pump start level [%], added pin
    fHiStop : REAL := 80.0;           // 停泵液位阈 [百分数]（可增引脚）/ Pump stop level [%], added pin
    tMinRun : TIME := T#30S;          // 最短运行时长 [毫秒] / Minimum run duration [ms]
    tMinOff : TIME := T#30S;          // 最短停机时长 [毫秒] / Minimum off duration [ms]
    tRunSwap: TIME := T#12H;          // 运行时长轮值阈 [毫秒] / Run-time swap threshold [ms]
    tHandover: TIME := T#10S;         // 交棒确认窗口 [毫秒] / Handover confirm window [ms]
END_VAR
VAR_OUTPUT
    bP1Req  : BOOL;                   // 泵 1 启动指令 / Pump 1 start command
    bP2Req  : BOOL;                   // 泵 2 启动指令 / Pump 2 start command
    bLead   : UINT;                   // 当前主泵号 [1 或 2] / Current lead pump [1 or 2]
    bError  : BOOL;                   // 故障标志，与故障级码配对（R45）/ Fault flag paired with fault codes
    uErrorId: UDINT;                  // 错误码，0 = 无错 / Error code, 0 = none
END_VAR
VAR
    rTrigSwap: R_TRIG;                // 手动轮换沿检测，每拍无条件刷新 / Manual swap edge detector
    tonMinRun: TON;                   // 最短运行计时，每拍无条件刷新 / Minimum run timer, refreshed every scan
    tonMinOff: TON;                   // 最短停机计时，每拍无条件刷新 / Minimum off timer, refreshed every scan
    tonRunTim: TON;                   // 主泵运行时长计时，每拍无条件刷新 / Lead run-time timer, refreshed every scan
    tonHandov: TON;                   // 交棒确认计时，每拍无条件刷新 / Handover confirm timer, refreshed every scan
    eState   : E_DL_TankPumpState;    // 内部状态机 / Internal state machine
    bLead1   : BOOL;                  // 主泵 1 标志 / Lead is pump 1 flag
    bLvlOk   : BOOL;                  // 液位输入有效 / Level input validity
    bStartReq: BOOL;                  // 液位低启泵请求 / Level-low start request
    bStopReq : BOOL;                  // 液位高停泵请求 / Level-high stop request
    bSwapReq : BOOL;                  // 本拍轮换请求 / Swap request this scan
    bBothFb  : BOOL;                  // 双泵反馈同时有效 / Both feedbacks valid
    bFbDualFail: BOOL;                // 双泵反馈双失效 / Both feedbacks failed
    bSwapWait: BOOL;                  // 交棒等待中 / Handover waiting flag
    bIntrlk  : BOOL;                  // 硬联锁激活 / Hard interlock active flag
END_VAR
VAR CONSTANT
    DL_TLC_FIN  : REAL := 1.0E30;     // REAL 有限幅值判界 / REAL finiteness magnitude bound
END_VAR

// ---- 段 1｜边沿与定时器实例无条件周期刷新（红线：禁入条件分支）----------------
rTrigSwap(CLK := bSwap);                              // 手动轮换沿检测 / Manual swap edge detection
tonMinRun(IN := (bP1Req OR bP2Req) AND (eState = eLeadRun), PT := tMinRun); // 最短运行计时 / Minimum run timing
tonMinOff(IN := (NOT (bP1Req OR bP2Req)) AND (eState = eIdle), PT := tMinOff); // 最短停机计时 / Minimum off timing
tonRunTim(IN := (eState = eLeadRun) AND (bP1Req OR bP2Req), PT := tRunSwap); // 运行时长轮值计时 / Run-time rotation timing
tonHandov(IN := bSwapWait, PT := tHandover);          // 交棒确认计时 / Handover confirm timing

// ---- 段 2｜输入有效性与回差判据 ------------------------------------------------
bLvlOk := (fLevel = fLevel) AND (ABS(fLevel) < DL_TLC_FIN); // 液位有限 / Level finite
bStartReq := bLvlOk AND (fLevel < fLoStart);          // 液位低于启泵阈 / Level below start threshold
bStopReq  := bLvlOk AND (fLevel > fHiStop);           // 液位高于停泵阈 / Level above stop threshold

// ---- 段 3｜状态机（CASE 带 ELSE 锁安全侧：双泵停）--------------------------------
CASE eState OF
    eIdle:
        bP1Req := FALSE;                              // 待机双泵停 / Both off in idle
        bP2Req := FALSE;                              // 待机双泵停 / Both off in idle
        IF bAuto AND bLvlOk AND bStartReq AND (NOT bLoLo) AND tonMinOff.Q THEN
            eState := eLeadRun;                       // 低液位且停机时满启主泵 / Level low and off-time met, start lead
        END_IF
    eLeadRun:
        IF bLead1 THEN
            bP1Req := bAuto AND (NOT bStopReq) AND (NOT bHiHi); // 主泵 1 指令 / Pump 1 command
            bP2Req := FALSE;                          // 备泵停 / Standby off
        ELSE
            bP2Req := bAuto AND (NOT bStopReq) AND (NOT bHiHi); // 主泵 2 指令 / Pump 2 command
            bP1Req := FALSE;                          // 备泵停 / Standby off
        END_IF
        bSwapReq := (tonRunTim.Q OR rTrigSwap.Q) AND bAuto AND bLvlOk; // 轮值时长满或手动沿请求轮换 / Rotation or manual swap request
        IF bSwapReq AND (NOT bHiHi) AND (NOT bLoLo) THEN
            IF bLead1 THEN
                bP2Req := TRUE;                       // 交棒先启新主泵（不断流时序）/ Handover starts new lead first
            ELSE
                bP1Req := TRUE;                       // 交棒先启新主泵 / Handover starts new lead first
            END_IF
            bSwapWait := TRUE;                        // 进入交棒等待 / Enter handover wait
            eState := eSwapWait;                      // 转交棒等待态 / To swap wait state
        ELSIF ((NOT bAuto) OR bStopReq OR (NOT bLvlOk)) AND tonMinRun.Q THEN
            bP1Req := FALSE;                          // 停泵条件且最短运行时满（防频启）/ Stop conditions with min-run met
            bP2Req := FALSE;                          // 停泵条件双停 / Stop conditions stop both
            IF (NOT bLvlOk) THEN
                uErrorId := 16#0005_00B2;             // 信息级：液位非有限冻结投切 / Info: non-finite freezes switching
            END_IF
            eState := eIdle;                          // 回待机 / Back to idle
        END_IF
    eSwapWait:
        bSwapWait := TRUE;                            // 等待标志保持 / Wait flag held
        IF bLead1 THEN
            bP1Req := TRUE;                           // 旧主泵保持运行 / Old lead kept running
            bP2Req := TRUE;                           // 新主泵等待反馈 / New lead awaiting feedback
            bBothFb := bP1Fb AND bP2Fb;               // 双反馈确认 / Both feedbacks confirmed
        ELSE
            bP2Req := TRUE;                           // 旧主泵保持运行 / Old lead kept running
            bP1Req := TRUE;                           // 新主泵等待反馈 / New lead awaiting feedback
            bBothFb := bP1Fb AND bP2Fb;               // 双反馈确认 / Both feedbacks confirmed
        END_IF
        IF bBothFb THEN
            IF bLead1 THEN
                bP1Req := FALSE;                      // 新主泵确认后停旧泵（停止侧安全执行）/ Stop old lead after confirm
                bLead1 := FALSE;                      // 轮值交棒完成 / Rotation handed over
            ELSE
                bP2Req := FALSE;                      // 新主泵确认后停旧泵 / Stop old lead after confirm
                bLead1 := TRUE;                       // 轮值交棒完成 / Rotation handed over
            END_IF
            bSwapWait := FALSE;                       // 清等待标志 / Clear wait flag
            eState := eLeadRun;                       // 回单主泵运行态 / Back to lead running
        ELSIF tonHandov.Q THEN
            IF bLead1 THEN
                bP2Req := FALSE;                      // 等待超时撤新泵请求撤轮换 / Timeout revokes new lead
            ELSE
                bP1Req := FALSE;                      // 等待超时撤新泵请求撤轮换 / Timeout revokes new lead
            END_IF
            bSwapWait := FALSE;                       // 清等待标志 / Clear wait flag
            eState := eLeadRun;                       // 回原主泵运行态 / Back to original lead
            uErrorId := 16#0005_00B2;                 // 信息级：交棒等待超时回落 / Info: handover wait timeout
        END_IF
    eFault:
        bP1Req := FALSE;                              // 故障态双泵停 / Both off in fault
        bP2Req := FALSE;                              // 故障态双泵停 / Both off in fault
        bSwapWait := FALSE;                           // 故障清等待 / Fault clears wait
        IF (NOT bP1Fb) AND (NOT bP2Fb) THEN
            eState := eIdle;                          // 可达解除路径：双泵实停复归 / Reachable release: both stopped
            uErrorId := 16#0000_0000;                 // 清码 / Clear code
        END_IF
    ELSE
        eState := eFault;                             // 非法状态兜底 / Illegal state fallback
END_CASE

// ---- 段 4｜双泵反馈双失效监视（运行指令下反馈缺失）------------------------------
bFbDualFail := (bP1Req AND NOT bP1Fb) AND (bP2Req AND NOT bP2Fb); // 双指令双无反馈 / Both commanded, both no feedback
IF bFbDualFail THEN
    eState := eFault;                                 // 双失效锁故障 / Dual failure latches fault
END_IF

// ---- 段 5｜HiHi/LoLo 独立硬联锁窗（直接切输出，不进状态机）----------------------
bIntrlk := bHiHi OR bLoLo;                            // 硬联锁激活判定 / Interlock active detection
IF bHiHi THEN
    bP1Req := FALSE;                                  // 高高位独立窗双泵停 / HiHi window stops both
    bP2Req := FALSE;                                  // 高高位独立窗双泵停 / HiHi window stops both
END_IF
IF bLoLo THEN
    bP1Req := TRUE;                                   // 低低位独立窗双泵启（恢复液位安全侧）/ LoLo window starts both
    bP2Req := TRUE;                                   // 低低位独立窗双泵启 / LoLo window starts both
END_IF

// ---- 段 6｜主泵号输出与错误码装配 ----------------------------------------------
IF bLead1 THEN
    bLead := 1;                                       // 主泵号输出 / Lead pump number output
ELSE
    bLead := 2;                                       // 主泵号输出 / Lead pump number output
END_IF
IF bIntrlk THEN
    bError   := TRUE;                                 // 硬联锁故障配对（R45）/ Interlock fault paired
    uErrorId := 16#0005_00B4;                         // 码位：硬联锁触发 / Code: hard interlock
ELSIF eState = eFault THEN
    bError   := TRUE;                                 // 双失效故障配对 / Dual failure fault paired
    uErrorId := 16#0005_00B3;                         // 码位：双泵失效 / Code: dual pump failure
ELSIF eState = eSwapWait THEN
    bError   := FALSE;                                // 信息级不置故障 / Info never sets fault
    uErrorId := 16#0005_00B2;                         // 信息级：交棒等待 / Info: handover wait
ELSE
    bError   := FALSE;                                // 无错清标志 / Clear fault flag
    uErrorId := 16#0000_0000;                         // 无码 / No code
END_IF
END_FUNCTION_BLOCK

(* ---- FB_DL_TankLevelStrapping.st ---- *)
(*
  FB_DL_TankLevelStrapping  —  储罐液位-容积分层标定与体积折算 / Tank level-volume strapping table conversion
  分类 Category : DL_Process
  码位 Code     : 16#06_0_BA
  段位说明      : R38 W7 预留 B6~BF 本轮正式启用，B9 格由 RadiatorZoneValve 启用，本件启用 BA 格
  版本 Version  : 1.0.0
  来源 Source   : 自研线（t2-1-lgf-math 次源）— 容积表标定核对待挖项
  溯源 Origin   : clean-room 实现，分层容积表折算为计量公开语义，未复制任何源码行
                  （与 FC_DL_MultiPointLinear 分工：那件是通用折算原子，本件带标定核对与罐型组态语义）
  功能 Function : 1) 分层容积表折算：液位 [m] → 体积 [m³]，走 FC_DL_MultiPointLinear 分段线性原子；
                  2) 越表插值拒绝：实测液位越出表界（外推被拒）时体积出口置 0 并置信息级码；
                  3) 标定核对：核对点（参考液位/参考体积）入容差窗（FB_DL_ToleranceWindow）判定，
                  核对失败锁故障（防表错继续计量），bReset 解除；
                  4) 液位百分比出口：FC_DL_LinearScale 表界归一。
  边界 Boundary : ① 表合法性（折点 >= 2 且液位严格递增）由折算原子校验，本件透传其错误码并锁存；
                  ② fTankMaxVolM3 为组态罐容上限：折算结果越上限钳制 + 信息级码（防表末段误配）；
                  ③ 组态域闸覆盖全部参与换算引脚（R151）；核对容差/参考体积域非法判组态错；
                  ④ 无状态机相（折算型 FB）：核对失败经锁存位承载，无跨相 TON 复用问题；
                  ⑤ R228-B 达标声明：eFault 迁出 = rtReset.Q（输入引脚，恒可达），逐字写于此；
                  ⑥ 折算原子为 LREAL 口径：入参/返回显式 REAL_TO_LREAL / LREAL_TO_REAL 转换。
  依赖 Depends  : FC_DL_MultiPointLinear / FC_DL_LinearScale（函数调用，引脚按 registry 实名）；
                  FB_DL_ToleranceWindow（实例化，引脚按 registry 实名）
  码表 Error codes（本件格 06_0_BA，子码步进 +0x100）:
    16#0006_01BA 信息级：标定核对通过（bCalCheck 拍）
    16#0006_02BA 故障级：标定核对失败（核对点越容差窗），锁存至复位
    16#0006_03BA 故障级：容积表非法（折点不足或非严格递增），锁存至复位
    16#0006_04BA 信息级：实测液位越表界，体积拒绝输出（置 0）
    16#0006_05BA 故障级：组态非法（点数/参考量/罐容上限域非法），锁存至复位
    16#0006_06BA 信息级：折算体积越组态罐容上限，已钳制
    16#0006_07BA 故障级：状态机落 ELSE 兜底（非法状态 ID）

  修订历史 Revision :
    2026-11-19  v1.0.0  R39 首版（批次 4 · 序号 18）
*)

TYPE E_DL_StrapState :
(
    eReady      := 0,    // 就绪：表合法且液位在表界内 / Ready, table valid and level in range
    eTableBad   := 10,   // 表非法：折算原子校验失败 / Table invalid, interpolator check failed
    eOutOfRange := 20,   // 越表：实测液位越表界 / Out of table range
    eCalFail    := 30,   // 核对失败：标定核对越容差 / Calibration check failed
    eFault      := 90    // 组态/核对故障锁定 / Fault, latched
);
END_TYPE

FUNCTION_BLOCK FB_DL_TankLevelStrapping
VAR_INPUT
    fLevelMeasM   : REAL := 0.0;         // 实测液位 [m] / Measured liquid level
    nTablePts     : INT := 0;            // 容积表有效折点数 [个]，2..16 / Strapping table point count
    fTankMaxVolM3 : REAL := 1000.0;      // 组态罐容上限 [m³]，域 > 0 / Tank volume configuration ceiling
    fRefLevelM    : REAL := 0.0;         // 核对点参考液位 [m] / Reference level for calibration check
    fRefVolM3     : REAL := 0.0;         // 核对点参考体积 [m³]，域 > 0 / Reference volume for check
    fRefTolPct    : REAL := 1.0;         // 核对容差 [%]（相对参考体积），域 (0, 100] / Check tolerance in percent
    bCalCheck     : BOOL := FALSE;       // 标定核对指令（上升沿）/ Calibration check command
    bReset        : BOOL := FALSE;       // 故障复位，上升沿生效 / Fault reset, rising edge
END_VAR
VAR_OUTPUT
    fVolumeM3    : REAL;                 // 折算体积 [m³]（越表/故障置 0）/ Converted volume output
    fLevelPct    : REAL;                 // 液位百分比 [%]（表界归一）/ Level percent of table span
    bOutOfRange  : BOOL;                 // 越表拒绝标志（瞬时，每拍重算）[-] / Out-of-range rejection flag
    bTableValid  : BOOL;                 // 容积表合法性 [-] / Table validity flag
    bCalOk       : BOOL;                 // 最近一次核对通过锁存 [-] / Last check passed latch
    eState       : E_DL_StrapState;      // 状态出口，段尾单点映射 / State outlet
    bError       : BOOL;                 // 故障锁存，仅故障级码置位，bReset 清除 [-] / Fault latch
    uErrorId     : UDINT;                // 事件码，0 = 无事件（故障级锁存回放）/ Event code
END_VAR
VAR_IN_OUT
    afLevelM : ARRAY[0..15] OF LREAL;    // 容积表液位折点 [m]，须严格递增 / Table level breakpoints, strictly increasing
    afVolM3  : ARRAY[0..15] OF LREAL;    // 容积表体积折点 [m³] / Table volume breakpoints
END_VAR
VAR
    fbTol      : FB_DL_ToleranceWindow;  // 核对容差窗实例（主体首部无条件刷新）/ Check tolerance window instance
    rtCalCheck : R_TRIG;                 // 核对指令上升沿 / Check command rising edge
    rtReset    : R_TRIG;                 // 复位上升沿 / Reset rising edge
    _lrVolCalc : LREAL;                  // 主折算体积中间量 [m³]（LREAL 口径）/ Main volume working value
    _lrVolAtRef: LREAL;                  // 核对点折算体积 [m³] / Volume at reference level
    _nSegMain  : INT;                    // 主折算命中段号 / Main conversion segment index
    _bExtrap   : BOOL;                   // 主折算外推标志 / Main conversion extrapolation flag
    _bClamp    : BOOL;                   // 主折算钳位标志 / Main conversion clamp flag
    _uMplErr   : UDINT;                  // 折算原子错误码透传 / Interpolator error passthrough
    _nSegRef   : INT;                    // 核对折算命中段号 / Check conversion segment index
    _bExtRef   : BOOL;                   // 核对折算外推标志 / Check conversion extrapolation flag
    _bClpRef   : BOOL;                   // 核对折算钳位标志 / Check conversion clamp flag
    _uErrRef   : UDINT;                  // 核对折算错误码透传 / Check conversion error passthrough
    _fScalePct : REAL;                   // 百分比中间量 [%] / Percent working value
    _bScaleOk  : BOOL;                   // 百分比换算有效 / Percent scaling valid
    _bTolSt    : BOOL;                   // 容差窗状态回传保持变量（有状态纪律）/ Tolerance window state hold member
    _bCalRun   : BOOL;                   // 本拍执行核对标志 / Check executed this cycle
    _eStateInt : E_DL_StrapState := E_DL_StrapState.eReady;   // 内部状态（CASE 唯一写入目标）/ Internal state
    _uInfo     : UDINT;                  // 信息码，每拍重算 / Info code
    _uFault    : UDINT;                  // 故障码锁存寄存 / Latched fault code register
    _bFault    : BOOL;                   // 故障锁存位 / Latched fault bit
    _bCfgBad   : BOOL;                   // 组态非法聚合 / Configuration invalid aggregate
END_VAR
VAR CONSTANT
    DL_TLS_INF_CAP  : REAL := 1.0E15;    // 非有限值筛查幅值上限 / Non-finite screening cap
    DL_TLS_PTS_MAX  : INT   := 16;       // 折点数上限（= 数组维度）/ Point count upper bound
    DL_TLS_VOL_EPS  : LREAL := 1.0E-9;   // 容差半宽下限兜底 [m³] / Tolerance half-width floor
END_VAR

(* —— 段 0：边沿实例无条件周期刷新（R182：调用语句不得置于 IF/CASE 内） —— *)
(* 容差窗 fbTol 在段 8 调用（数据流：核对折算先于判定），仍为顶层无条件调用 *)
rtCalCheck(CLK := bCalCheck);                            // 核对沿刷新，每拍必调
rtReset(CLK := bReset);                                  // 复位沿刷新，每拍必调

(* —— 段 1：单拍量预清零（锁存量 _uFault/_bFault/bCalOk 不入清单，R187①） —— *)
_uInfo := 16#0000_0000;             // 信息码每拍重算
_bCfgBad := FALSE;                  // 组态非法预清零
bOutOfRange := FALSE;               // 越表标志缺省 FALSE（段 4 单点置位）
uErrorId := 16#0000_0000;           // 事件码缺省无事件

(* —— 段 2：组态域闸（覆盖全部参与判据换算的引脚，R151） —— *)
IF (nTablePts < 2) OR (nTablePts > DL_TLS_PTS_MAX) THEN
    _bCfgBad := TRUE;               // 折点数域非法
END_IF
IF (fTankMaxVolM3 <= 0.0) OR (ABS(fTankMaxVolM3) > DL_TLS_INF_CAP)
   OR (fRefVolM3 <= 0.0) OR (ABS(fRefVolM3) > DL_TLS_INF_CAP)
   OR (fRefTolPct <= 0.0) OR (fRefTolPct > 100.0)
   OR (fLevelMeasM <> fLevelMeasM) OR (ABS(fLevelMeasM) > DL_TLS_INF_CAP) OR ((fLevelMeasM - fLevelMeasM) <> 0.0) THEN
    _bCfgBad := TRUE;               // 罐容/参考量/容差/液位域非法
END_IF

(* —— 段 3：故障锁存与迁出沿（R228-B：rtReset.Q 恒可达） —— *)
IF _bCfgBad AND (NOT _bFault) THEN
    _uFault := 16#0006_05BA;        // 故障级：组态非法（仅首次进入时写入）
    _bFault := TRUE;
END_IF
IF rtReset.Q AND (NOT _bCfgBad) THEN
    _bFault := FALSE;               // 清故障锁存位（组态恢复合法为前提）
    _uFault := 16#0000_0000;
    bCalOk := FALSE;                // 核对通过锁存随复位清除
END_IF

(* —— 段 4：主折算（FC_DL_MultiPointLinear 原子；bClamp = FALSE，越表由外推标志承载拒绝语义） —— *)
_lrVolCalc := FC_DL_MultiPointLinear(afX := afLevelM,        // 液位折点表
                                     afY := afVolM3,         // 体积折点表
                                     fIn := REAL_TO_LREAL(fLevelMeasM),   // 实测液位（显式升型）
                                     nCount := nTablePts,    // 有效折点数
                                     bClamp := FALSE,        // 不钳位：越表拒绝语义自管
                                     nSegment => _nSegMain,  // 命中段号
                                     bExtrapolated => _bExtrap,   // 外推标志
                                     bClamped => _bClamp,    // 钳位标志
                                     uErrorId => _uMplErr);  // 错误码透传
bTableValid := (_uMplErr = 0) AND (_nSegMain >= 0);          // 表合法 = 无错误码且命中段有效

(* —— 段 5：液位百分比出口（FC_DL_LinearScale 原子，表界归一；表非法时出口 0） —— *)
IF bTableValid THEN
    _fScalePct := FC_DL_LinearScale(fIn := fLevelMeasM,      // 实测液位
                                    fInMin := LREAL_TO_REAL(afLevelM[0]),       // 表界下端
                                    fInMax := LREAL_TO_REAL(afLevelM[nTablePts - 1]),   // 表界上端（下标已由点数闸钳位）
                                    fOutMin := 0.0,          // 归一 0%
                                    fOutMax := 100.0,        // 归一 100%
                                    bClamp := TRUE,          // 表界内归一，越界钳位
                                    bValid => _bScaleOk,     // 换算有效标志
                                    uErrorId => _uInfo);     // 换算错误码（瞬时，并入信息码）
ELSE
    _fScalePct := 0.0;               // 表非法：百分比出口置 0（防御口径）
END_IF
fLevelPct := _fScalePct;            // 百分比出口镜像

(* —— 段 6：状态分类 CASE（计算型分类，含 ELSE 兜底） —— *)
CASE _eStateInt OF

E_DL_StrapState.eReady:
    IF _bFault THEN
        _eStateInt := E_DL_StrapState.eFault;           // 故障锁存：进故障态
    ELSIF NOT bTableValid THEN
        _eStateInt := E_DL_StrapState.eTableBad;        // 表非法：进表错态
    ELSIF _bExtrap THEN
        _eStateInt := E_DL_StrapState.eOutOfRange;      // 越表：进拒绝态
    END_IF

E_DL_StrapState.eTableBad:
    IF bTableValid THEN
        _eStateInt := E_DL_StrapState.eReady;           // 表恢复合法：回就绪态
    END_IF

E_DL_StrapState.eOutOfRange:
    IF (NOT _bExtrap) AND bTableValid THEN
        _eStateInt := E_DL_StrapState.eReady;           // 回表界内：回就绪态
    END_IF

E_DL_StrapState.eCalFail:
    IF (NOT _bFault) AND bTableValid THEN
        _eStateInt := E_DL_StrapState.eReady;           // 核对故障解除：回就绪态
    END_IF

E_DL_StrapState.eFault:
    IF NOT _bFault THEN
        _eStateInt := E_DL_StrapState.eReady;           // 故障解除：回就绪态
    END_IF

ELSE
    _uFault := 16#0006_07BA;        // 故障级：非法状态 ID 兜底
    _bFault := TRUE;
    _eStateInt := E_DL_StrapState.eFault;   // 强制回故障态

END_CASE

(* —— 段 7：体积出口合成（越表拒绝 / 表非法 / 故障三路置 0；越罐容上限钳制） —— *)
IF _bFault OR (NOT bTableValid) OR _bExtrap THEN
    IF _bExtrap AND (NOT _bFault) AND bTableValid THEN
        bOutOfRange := TRUE;        // 越表拒绝标志（瞬时）
        _uInfo := 16#0006_04BA;     // 信息级：越表拒绝输出
    END_IF
    IF (NOT bTableValid) AND (NOT _bFault) THEN
        _uFault := 16#0006_03BA;    // 故障级：容积表非法（锁存）
        _bFault := TRUE;
    END_IF
    fVolumeM3 := 0.0;               // 拒绝/非法/故障：体积出口置 0
ELSE
    IF _lrVolCalc > REAL_TO_LREAL(fTankMaxVolM3) THEN
        fVolumeM3 := fTankMaxVolM3; // 越罐容上限钳制
        _uInfo := 16#0006_06BA;     // 信息级：已钳制
    ELSE
        fVolumeM3 := LREAL_TO_REAL(_lrVolCalc);     // 正常折算出口（显式降型）
    END_IF
END_IF

(* —— 段 8：标定核对（沿触发核对折算 → fbTol 顶层判定 → 自消费判定标志） —— *)
IF rtCalCheck.Q AND (NOT _bFault) AND bTableValid THEN
    _lrVolAtRef := FC_DL_MultiPointLinear(afX := afLevelM,      // 液位折点表
                                          afY := afVolM3,       // 体积折点表
                                          fIn := REAL_TO_LREAL(fRefLevelM),     // 核对点参考液位
                                          nCount := nTablePts,  // 有效折点数
                                          bClamp := FALSE,      // 不钳位
                                          nSegment => _nSegRef, // 命中段号
                                          bExtrapolated => _bExtRef,    // 外推标志
                                          bClamped => _bClpRef, // 钳位标志
                                          uErrorId => _uErrRef);    // 错误码透传
    IF (_uErrRef = 0) AND (_nSegRef >= 0) AND (NOT _bExtRef) THEN
        _bCalRun := TRUE;           // 核对折算有效：判定标志置位（本段末尾自消费）
        _eStateInt := E_DL_StrapState.eCalFail;     // 判定期间暂入核对态（按结果迁出）
    ELSE
        _uFault := 16#0006_02BA;    // 故障级：核对点越表（核对失败口径之一）
        _bFault := TRUE;
    END_IF
END_IF
fbTol(bEnable := _bCalRun,                               // 仅核对拍判定
      fTarget := REAL_TO_LREAL(fRefVolM3),               // 核对目标体积
      fActual := _lrVolAtRef,                            // 核对点折算体积
      fTolerance := MAX(REAL_TO_LREAL(fRefVolM3) * REAL_TO_LREAL(fRefTolPct) / 100.0, DL_TLS_VOL_EPS),   // 容差半宽（相对口径，下限防零窗死判）
      fHysteresis := 0.0);                               // 无回差（单次判定口径）
IF _bCalRun THEN
    IF fbTol.bOk THEN
        bCalOk := TRUE;             // 核对通过锁存
        _uInfo := 16#0006_01BA;     // 信息级：核对通过
        _eStateInt := E_DL_StrapState.eReady;   // 回就绪态
    ELSE
        _uFault := 16#0006_02BA;    // 故障级：标定核对失败（锁存至复位）
        _bFault := TRUE;
    END_IF
    _bCalRun := FALSE;              // 判定标志自消费（单拍口径）
END_IF

(* —— 段 9：出口单点映射（名实同源；锁存码回放，禁同拍抹除） —— *)
IF _bFault THEN
    uErrorId := _uFault;            // 故障锁存码回放（不在故障态按当下输入重推）
    bError := TRUE;
    bOutOfRange := FALSE;           // 故障态越表标志强制 FALSE（口径归一）
ELSE
    uErrorId := _uInfo;             // 信息码
    bError := FALSE;
END_IF
eState := _eStateInt;               // 状态出口单点映射

END_FUNCTION_BLOCK

(* ---- FB_DL_TempCompClassify.st ---- *)
(*==============================================================================
 * 组件名称 (Component)  : FB_DL_TempCompClassify
 * 所属子库 (Sublibrary) : DL_Process
 * 当前版本 (Version)    : 1.0.0
 * 兼容性   (Platform)   : CODESYS 3.5+ / TwinCAT 3 / 汇川 InoProShop / 施耐德 Machine Expert
 *                         仅依赖 Standard.library（R_TRIG），零厂商私有库
 * 功能描述 (Function)   : 组件功率温度补偿分档。
 *                         把实测功率按温度系数归一到一个基准温度，再把归一功率切成四档（G1 最低 … G4 最高），
 *                         相邻档之间带迟滞带，防止测点在分界线上抖动造成档位来回跳。
 *                         归一式（百分比系数口径，写死）：
 *                           P_norm = P_meas · (1 + k/100 · (T_meas − T_ref))
 *                           k 单位 %/°C，正 k 表示"温度升高时实测功率升高"，归一化需回减；
 *                           该式在 k/100·ΔT ≤ −1 时会出现非正比例因子，此时判 eNormCollapse 并停判。
 *                         分档结构（三阈值四档，迟滞带 fHyst 双向对称）：
 *                           升档：P_norm > fThN + fHyst 才升到 N+1
 *                           降档：P_norm < fThN − fHyst 才降到 N
 *                           带内（含边界）保持当前档 —— 这就是迟滞的全部作用，无其它隐藏状态。
 *                         验收向量：
 *                           ① k=0 之外的正常参数：P=1000 W, T=35 °C, k=+2 %/°C, Tref=25 °C
 *                              → 比例因子 1+0.02×10 = 1.20，P_norm = 1200 W
 *                           ② 阈值 800/1000/1200 W，迟滞 20 W：P_norm=1210 且当前 G3 → 升 G4
 *                           ③ 同参 P_norm=1190 且当前 G4 → 保持 G4（未破 1200−20）
 *                           ④ 同参 P_norm=1170 且当前 G4 → 降 G3
 * 接口     (Interface)  : 入 bEnable 使能、fPowerMeas 实测功率、fTempMeas 实测温度、fTempCoeff 温度系数、
 *                         fTempRefC 基准温度、fTh1..fTh3 三阈值、fHyst 迟滞半宽、bReset 复位沿；
 *                         出 fPwrNorm 归一功率、iGrade 档位（1..4，0 = 未分级）、bValid 有效、
 *                         bGradeChanged 换档脉冲（单拍）、eState 相、eCause 成因、bError 故障标志。
 * 边界     (Boundary)   : ① **属主边界（写死）：本件只做"归一 + 分档"，不裁决组件是否合格、
 *                         不驱动负载功率设定**（属功率控制件）；② **温补系数零闸**：k = 0 或非有限
 *                         → 温补形同虚设且无任何可观测差异，属静默失效（R179），按故障级锁存；
 *                         ③ **阈值单调闸**：fTh1 < fTh2 < fTh3 且 fHyst ≥ 0，违反即锁存 eCfgIllegal；
 *                         ④ **迟滞半宽闸**：fHyst 必须小于最小相邻阈值间距的一半，否则档位可同时
 *                         满足升/降条件，出现"抖到死"或"跨档跳"，判 eCfgIllegal；
 *                         ⑤ **归一塌陷闸**：比例因子 ≤ 0 → 判 eNormCollapse（当拍不判档、bValid=FALSE，
 *                         不锁存，属样本侧异常而非组态异常）；
 *                         ⑥ 浮点比较一律用显式不等号 + 差值容差判等，禁 = / <> 直接判值；
 *                         ⑦ eFault 可迁出：bReset 上升沿 → eIdle，解除式恒可达（外部引脚门控）；
 *                         ⑧ 零全局耦合、零物理地址。
 * 分工声明 (Scope)      : 本件只管"功率温补与四档分级"。不接管：OCV 温度归一判带
 *                         （属 FB_DL_OcvTempNormalize）、温度闭环控制（属温控件）、
 *                         功率设定值下发（属功率环件）。
 * 来源标签 (Source Tag) : ROADMAP 空勾真缺口 P1（功率温补分档，自研 clean-room）
 * 码表     (Codes)      : 本件不占用任何全局数字码位（零码位范式 R297）；诊断由 BOOL + ENUM 出口承担。
 * 红线自检 (Redline)    : R1 ✓ 零 GVL/VAR_EXTERNAL ｜ R2 ✓ 零 %I/%Q/%M ｜ R3 ✓ 纯 IEC 61131-3
 *                         R4 ✓ 零闸 + 单调闸 + 迟滞配比闸 + 塌陷闸 + 容差 ｜ R5 ✓ 声明逐行同行双语注释
 *                         R6 ✓ ENUM+CASE 含 ELSE 兜底 ｜ R7 ✓ R_TRIG 段 0 无条件刷新（本件无 TON）
 * 修订历史 (Revision)   : 2026-11-19  v1.0.0  R47 首版（批次 2 · 序号 8）
 *==============================================================================*)

TYPE E_DL_TccState :
(
    eIdle  := 0,    // 待机相（未使能） / Idle, disabled
    eRun   := 10,   // 分档相（归一与迟滞判档） / Running, normalise and classify
    eFault := 90    // 故障相（等复位） / Fault, awaiting reset
);
END_TYPE

TYPE E_DL_TccCause :
(
    eNone         := 0,   // 无异常 / No anomaly
    eCfgIllegal   := 1,   // 组态非法（阈值非单调 / 迟滞过宽） / Illegal configuration
    eCoeffZero    := 2,   // 温补系数为零或非有限（静默失效，故障级） / Zero or non-finite coefficient
    eNormCollapse := 3,   // 归一比例因子非正（样本侧异常，当拍不判） / Non-positive normalisation factor
    eSampleBad    := 4,   // 样本非有限（当拍不判） / Non-finite sample
    ePhaseBad     := 5    // 非法相位兜底 / Illegal phase fallback
);
END_TYPE

FUNCTION_BLOCK FB_DL_TempCompClassify
VAR_INPUT
    bEnable    : BOOL := FALSE;      // 使能（FALSE 冻结分档） [-] / Enable
    fPowerMeas : LREAL := 0.0;       // 实测功率 [W] / Measured power [W]
    fTempMeas  : LREAL := 25.0;      // 实测温度 [°C] / Measured temperature [°C]
    fTempCoeff : LREAL := 2.0;       // 温度系数，域 ≠ 0 且有限 [%/°C] / Temperature coefficient, non-zero and finite
    fTempRefC  : LREAL := 25.0;      // 基准温度 [°C] / Reference temperature [°C]
    fTh1       : LREAL := 800.0;     // 一档/二档分界 [W] / G1-G2 boundary [W]
    fTh2       : LREAL := 1000.0;    // 二档/三档分界 [W] / G2-G3 boundary [W]
    fTh3       : LREAL := 1200.0;    // 三档/四档分界 [W] / G3-G4 boundary [W]
    fHyst      : LREAL := 20.0;      // 迟滞半宽（对称），域 ≥ 0 [W] / Symmetric hysteresis half-width, >= 0
    bReset     : BOOL := FALSE;      // 故障复位沿 [-] / Fault reset edge
END_VAR
VAR_OUTPUT
    fPwrNorm      : LREAL := 0.0;                        // 归一到基准温度后的功率 [W] / Power normalised to the reference temperature
    iGrade        : INT := 0;                            // 档位 1..4（0 = 未分级） [档] / Grade 1..4, 0 = ungraded
    bValid        : BOOL := FALSE;                       // 结果有效 [-] / Result valid
    bGradeChanged : BOOL := FALSE;                       // 换档脉冲（单拍） [-] / Grade-change pulse, single scan
    eState        : E_DL_TccState := E_DL_TccState.eIdle;   // 相出口 [-] / Phase outlet
    eCause        : E_DL_TccCause := E_DL_TccCause.eNone;   // 成因出口（R190 归因唯一） [-] / Cause outlet
    bError        : BOOL := FALSE;                       // 故障标志（仅故障级成因） [-] / Error flag, fault level only
END_VAR
VAR
    _eState   : E_DL_TccState := E_DL_TccState.eIdle;    // 内部相（CASE 唯一写入目标） / Internal phase
    _eCause   : E_DL_TccCause := E_DL_TccCause.eNone;    // 成因锁存量 / Latched cause
    _bFault   : BOOL := FALSE;                           // 故障锁存位 / Latched fault bit
    _iGrade   : INT := 0;                                // 内部档位（迟滞保持量） / Internal grade, hysteresis state
    _fNorm    : LREAL := 0.0;                            // 归一功率工作值 [W] / Normalised power working value
    _fRatio   : LREAL := 0.0;                            // 归一比例因子 [-] / Normalisation ratio
    _bChanged : BOOL := FALSE;                           // 换档脉冲内部位（单拍） / Internal grade-change pulse
    _bCfgBad  : BOOL := FALSE;                           // 组态非法当拍量 / Illegal configuration this scan
    _bSampleOk: BOOL := FALSE;                           // 样本有限性结论 / Sample finiteness result
    rtReset   : R_TRIG;                                  // 复位沿实例，段 0 无条件调用 / Reset edge instance
END_VAR
VAR CONSTANT
    DL_TCC_EPS  : LREAL := 1.0E-9;   // 浮点判等容差（仅"贴边界"判定） [W] / Equality tolerance
    DL_TCC_PCT  : LREAL := 100.0;    // 百分数换算因子 [%] / Percentage scaling factor
    DL_TCC_WMIN : LREAL := 0.0;      // 归一功率下界（功率不许为负） [W] / Lower bound of the normalised power
END_VAR

(* —— 段 0：两沿无条件周期刷新（R228A；本件无 TON） —— *)
rtReset(CLK := bReset);                                          // 复位沿 / Reset edge

(* —— 段 1：单拍/输出量预置（锁存量 _eCause/_bFault/_iGrade 不入清单，R107） —— *)
fPwrNorm      := 0.0;                                            // 归一功率预置 / Normalised power preset
iGrade        := 0;                                              // 档位预置为未分级 / Grade preset to ungraded
bValid        := FALSE;                                          // 有效位预置 / Validity preset
_bChanged     := FALSE;                                          // 换档脉冲预清 / Grade-change pulse preset
bError        := FALSE;                                          // 故障标志预清（R45 配对） / Error preset
_fNorm        := 0.0;                                            // 工作值预置 / Working value preset
_fRatio       := 0.0;                                            // 比例因子预置 / Ratio preset

(* —— 段 2：组态闸（阈值单调 / 迟滞非负 / 迟滞不吞掉最窄间距） —— *)
_bCfgBad := NOT ((fTh1 < fTh2) AND (fTh2 < fTh3))                // 三阈值须严格单调 / Thresholds strictly monotonic
        OR (fHyst < 0.0)                                         // 迟滞半宽须非负 / Hysteresis must be non-negative
        OR (fHyst > ((fTh2 - fTh1) / 2.0))                       // 迟滞须小于最窄间距的一半 / Below half the narrowest gap
        OR (fHyst > ((fTh3 - fTh2) / 2.0));                      // 迟滞须小于最窄间距的一半（另一段同源约束） / Same constraint on the other gap
IF _bCfgBad THEN
    _eCause := E_DL_TccCause.eCfgIllegal;                        // 归因：组态非法 / Cause: illegal configuration
    _bFault := TRUE;                                             // 锁存 / Latch
    _eState := E_DL_TccState.eFault;                             // 入故障相 / Enter fault phase
END_IF

(* —— 段 3：温补系数零闸（k=0 使归一恒等，静默失效，故障级 R179） —— *)
IF (_eState <> E_DL_TccState.eFault) THEN
    IF (fTempCoeff = 0.0) OR (fTempCoeff <> fTempCoeff) OR ((fTempCoeff - fTempCoeff) <> (fTempCoeff - fTempCoeff)) THEN
        _eCause := E_DL_TccCause.eCoeffZero;                     // 归因：系数为零或非有限 / Cause: zero or non-finite coefficient
        _bFault := TRUE;                                         // 锁存 / Latch
        _eState := E_DL_TccState.eFault;                         // 入故障相 / Enter fault phase
    END_IF
END_IF

(* —— 段 4：迁出链（bReset 上升沿 → 待机相，并清档位保持量） —— *)
IF rtReset.Q THEN
    _bFault := FALSE;                                            // 清故障锁存 / Clear fault latch
    _eCause := E_DL_TccCause.eNone;                              // 清成因 / Clear cause
    _iGrade := 0;                                                // 档位保持量清零（复位后重新起档） / Grade cleared, restart classification
    _eState := E_DL_TccState.eIdle;                              // 回待机相 / Back to idle
END_IF

(* —— 段 5：相迁移（使能驱动；故障相由段 4 迁出） —— *)
CASE _eState OF

E_DL_TccState.eIdle:
    IF bEnable THEN
        _eState := E_DL_TccState.eRun;                           // 使能即进分档相 / Enable enters the running phase
    END_IF

E_DL_TccState.eRun:
    IF NOT bEnable THEN
        _eState := E_DL_TccState.eIdle;                          // 失能回待机相（不借故障相过桥，R211） / Disable returns to idle
    END_IF

E_DL_TccState.eFault:
    ;                                                            // 故障相：由段 4 复位沿迁出 / Exit handled by the reset edge

ELSE
    _eCause := E_DL_TccCause.ePhaseBad;                          // 归因：非法相位 / Cause: illegal phase
    _bFault := TRUE;                                             // 锁存 / Latch
    _eState := E_DL_TccState.eFault;                             // 强拉故障相 / Force fault phase

END_CASE

(* —— 段 6：归一（样本有限性 → 比例因子 → 归一功率，非有限当拍不判） —— *)
IF _eState = E_DL_TccState.eRun THEN
    _bSampleOk := NOT ((fPowerMeas <> fPowerMeas) OR ((fPowerMeas - fPowerMeas) <> (fPowerMeas - fPowerMeas)))
              AND NOT ((fTempMeas <> fTempMeas) OR ((fTempMeas - fTempMeas) <> (fTempMeas - fTempMeas)))
              AND NOT ((fTempRefC <> fTempRefC) OR ((fTempRefC - fTempRefC) <> (fTempRefC - fTempRefC)));
    IF _bSampleOk THEN
        _fRatio := 1.0 + ((fTempCoeff / DL_TCC_PCT) * (fTempMeas - fTempRefC));   // 归一比例因子 / Normalisation ratio
        IF _fRatio <= 0.0 THEN
            _eCause := E_DL_TccCause.eNormCollapse;              // 归因：比例因子非正（样本侧异常） / Cause: non-positive ratio
        ELSE
            _fNorm := fPowerMeas * _fRatio;                      // 归一功率 / Normalised power
            IF _fNorm < DL_TCC_WMIN THEN
                _fNorm := DL_TCC_WMIN;                           // 下钳（功率不许为负） / Clamp to the physical lower bound
            END_IF
            bValid := TRUE;                                      // 结果有效 / Result valid

            (* 四档迟滞判档：以内部保持量 _iGrade 为中心，只判"升一档/降一档/保持" *)
            CASE _iGrade OF
            0:                                                       // 未起档：按当前值定初始档（无迟滞，首次定向） / Initial assignment without hysteresis
                IF _fNorm > fTh3 THEN
                    _iGrade := 4;
                ELSIF _fNorm > fTh2 THEN
                    _iGrade := 3;
                ELSIF _fNorm > fTh1 THEN
                    _iGrade := 2;
                ELSE
                    _iGrade := 1;
                END_IF
                _bChanged := TRUE;                                   // 首次定档亦视为换档 / Initial assignment counts as a change

            1:
                IF _fNorm > (fTh1 + fHyst) THEN
                    _iGrade := 2;                                    // 升档（破上界 + 迟滞） / Step up
                    _bChanged := TRUE;
                END_IF

            2:
                IF _fNorm > (fTh2 + fHyst) THEN
                    _iGrade := 3;                                    // 升档 / Step up
                    _bChanged := TRUE;
                ELSIF _fNorm < (fTh1 - fHyst) THEN
                    _iGrade := 1;                                    // 降档（破下界 − 迟滞） / Step down
                    _bChanged := TRUE;
                END_IF

            3:
                IF _fNorm > (fTh3 + fHyst) THEN
                    _iGrade := 4;                                    // 升档 / Step up
                    _bChanged := TRUE;
                ELSIF _fNorm < (fTh2 - fHyst) THEN
                    _iGrade := 2;                                    // 降档 / Step down
                    _bChanged := TRUE;
                END_IF

            4:
                IF _fNorm < (fTh3 - fHyst) THEN
                    _iGrade := 3;                                    // 降档 / Step down
                    _bChanged := TRUE;
                END_IF

            ELSE
                _iGrade := 0;                                        // 档位保持量非法：归零重起（不锁存，属内部自愈） / Internal self-heal
            END_CASE

            iGrade := _iGrade;                                       // 档位出口（与本拍判定同源） / Grade outlet, same origin
        END_IF
    ELSE
        _eCause := E_DL_TccCause.eSampleBad;                         // 归因：样本非有限（当拍不判） / Cause: non-finite sample
    END_IF
END_IF

(* —— 段 7：出口单点映射（名实双出口，R191） —— *)
fPwrNorm      := _fNorm;                                             // 归一功率出口 / Normalised power outlet
bGradeChanged := _bChanged;                                          // 换档脉冲出口 / Grade-change outlet
eState        := _eState;                                            // 相出口 / Phase outlet
eCause        := _eCause;                                            // 成因出口 / Cause outlet
bError        := _bFault;                                            // 故障标志 / Error flag

END_FUNCTION_BLOCK

(* ---- FB_DL_TerminalReheatSeq.st ---- *)
(*
  FB_DL_TerminalReheatSeq  —  末端再热级联联锁 / Terminal reheat cascade interlock
  分类 Category : DL_Process
  码位 Code     : 16#06_0_B2
  版本 Version  : 1.0.0
  来源 Source   : t1-2-oscat-building — IEC 61131-3 标准语义的道莅防御性实现
  溯源 Origin   : clean-room 实现，VAV 再热级联公开控制语义借鉴，未复制任何源码行（RESUME 承接 R36 §4 #17 规格）
                  （级间延时语义对齐 FB_DL_SignalDebounce；变化率限幅对齐 FB_DL_RateLimiter，均不实例化）
  功能 Function : 1) 区域温度低于设定值产生再热需求，再热输出按级步进（级间延时 tStageDelay，防级联抖动）；
                  2) 风量低于 fMinAirflowPct 时再热按级降档（每 tStageDelay 降一级）并置 bMinAirflowLimit；
                  3) bReheatInhibit（制冷季互锁输入）时再热全关，出口镜像 bReheatInhibitActive；
                  4) 信号质量坏 → 保持当前级并置码（不跳变，规格强制）。
  边界 Boundary : ① fMinAirflowPct >= 100 判组态错（将使再热永久抑制）；fReheatStageStepPct <= 0 防除零判组态错；
                  ② 级数计算 nStage = TRUNC(fReheatCmdPct / fReheatStageStepPct) 后按级数上限钳制
                     （R28-2 两点向量：整除点 TRUNC 精确取整不越级；上限 +1 级钳到 fReheatMaxPct 对应级数不越上界）；
                  ③ 温度/风量信号非有限（NaN 用 x<>x 自反）→ 保持当前级并置码（不跳变）；
                  ④ 再热输出钳 [0, fReheatMaxPct]，禁越上限；
                  ⑤ 本件无状态机 ENUM/CASE（级联调节件），判据均为每拍重算或保持量承载，无锁存码。
  依赖 Depends  : 仅 Standard.library（TON/ABS/TRUNC/MIN/MAX）；语义对齐 FB_DL_RateLimiter / FB_DL_SignalDebounce（已注册）
  码表 Error codes（本件格 06_0_B2，子码步进 +0x100）:
    16#0006_01B2 信息级：信号质量坏（温度/风量非有限或越域），保持当前级
    16#0006_02B2 故障级：组态非法（最小风量 >= 100 / 级步 <= 0 / 上限越域）
    16#0006_03B2 信息级：最小风量约束生效（按级降档）
    16#0006_04B2 信息级：再热互锁生效，输出全关

  修订历史 Revision :
    2026-11-18  v1.0.0  R38 首版
*)

FUNCTION_BLOCK FB_DL_TerminalReheatSeq
VAR_INPUT
    fZoneTempC        : REAL := 22.0;     // 区域温度 [°C] / Zone temperature
    fZoneSetC         : REAL := 21.0;     // 区域设定值 [°C] / Zone setpoint
    fAirflowPct       : REAL := 80.0;     // 风量 [%] / Airflow percentage
    fMinAirflowPct    : REAL := 30.0;     // 最小风量 [%]，域 < 100 / Minimum airflow
    fReheatMaxPct     : REAL := 100.0;    // 再热上限 [%]，域 0..100 / Reheat ceiling
    fReheatStageStepPct: REAL := 20.0;    // 再热级步 [%]，域 > 0 / Reheat stage step
    tStageDelay       : TIME := T#10S;    // 级间延时 [ms]，域 > 0 / Stage change delay
    bReheatInhibit    : BOOL := FALSE;    // 再热互锁输入（制冷季）/ Reheat inhibit interlock input
END_VAR
VAR_OUTPUT
    fReheatCmdPct      : REAL;            // 再热输出指令 [%] / Reheat command
    bMinAirflowLimit   : BOOL;            // 最小风量约束生效 / Minimum airflow limit flag
    bReheatInhibitActive: BOOL;           // 互锁生效镜像出口（输入 bReheatInhibit 承载规格名）/ Inhibit active mirror
    nActiveStage       : INT;             // 当前再热级数 [级] / Active stage count
    nErrId             : UDINT;           // 事件码，0 = 无事件 / Event code
END_VAR
VAR
    tonStageDly : TON;                   // 级间延时计时（变化节流），自复位承载 / Stage change delay timer
    tonFaultWch : TON;                   // 故障观察窗，自复位 / Fault watch window, self-resetting
    _nStage     : INT;                   // 当前级数内部量 [级] / Internal stage count
    _nStageDes  : INT;                   // 期望级数（按需求算得）[级] / Desired stage count
    _nStageMax  : INT;                   // 级数上限 [级] / Stage ceiling
    _rErr       : REAL;                  // 温度偏差暂存 [K] / Temperature deviation scratch
    _bSigBad    : BOOL;                  // 信号质量坏聚合 / Signal quality bad aggregate
    _bStageBrk  : BOOL;                  // 级间延时窗断输入请求（自复位范式）/ Stage delay break request
    _bLimitHold : BOOL;                  // 最小风量约束保持量 / Airflow limit held quantity
    _uInfo      : UDINT;                 // 信息码，每拍重算 / Info code
    _bCfgBad    : BOOL;                  // 组态非法聚合 / Configuration invalid aggregate
END_VAR
VAR CONSTANT
    DL_WATCH_PT : TIME := T#2S;   // 故障观察窗 [ms]，自复位 / Fault watch window
END_VAR

(* —— 段 0：定时器无条件周期刷新（R182：调用语句不得置于 IF/CASE 内） —— *)
tonFaultWch(IN := (NOT tonFaultWch.Q), PT := DL_WATCH_PT);       // 观察窗自复位（表达式入参）
tonStageDly(IN := (NOT tonStageDly.Q) AND (NOT _bStageBrk), PT := tStageDelay);   // 级间延时自复位窗（表达式入参）
_bStageBrk := FALSE;                 // 断输入拍在调用后自清（R188 范式）

(* —— 段 1：单拍量预清零（保持量 _nStage/_bLimitHold 不入清单，R187①） —— *)
_uInfo := 16#0000_0000;              // 信息码每拍重算
bMinAirflowLimit := FALSE;           // 约束出口缺省 FALSE（段 6 单点置位）
_bCfgBad := FALSE;                   // 组态非法预清零
_bSigBad := FALSE;                   // 信号质量坏预清零
nErrId := 16#0000_0000;              // 事件码缺省无事件

(* —— 段 2：组态域闸（覆盖全部参与判据换算的引脚，R151） —— *)
IF fMinAirflowPct >= 100.0 THEN
    _bCfgBad := TRUE;                // 最小风量 >= 100：再热将永久抑制（规格强制）
END_IF
IF (fReheatStageStepPct <= 0.0) OR (fReheatStageStepPct <> fReheatStageStepPct) THEN
    _bCfgBad := TRUE;                // 级步非法（防除零）
END_IF
IF (fReheatMaxPct <= 0.0) OR (fReheatMaxPct > 100.0) OR (TIME_TO_DINT(tStageDelay) <= 0) THEN
    _bCfgBad := TRUE;                // 上限/级间延时非法
END_IF

(* —— 段 3：信号质量闸（温度/风量非有限或越域 → 保持当前级，不跳变） —— *)
IF (fZoneTempC <> fZoneTempC) OR (fZoneSetC <> fZoneSetC)
   OR (ABS(fZoneTempC) > 80.0) OR (ABS(fZoneSetC) > 80.0) THEN
    _bSigBad := TRUE;                // 温度信号质量坏
    _uInfo := 16#0006_01B2;          // 信息级：保持当前级
END_IF
IF (fAirflowPct <> fAirflowPct) OR (fAirflowPct < 0.0) OR (fAirflowPct > 150.0) THEN
    _bSigBad := TRUE;                // 风量信号质量坏
    _uInfo := 16#0006_01B2;          // 信息级：保持当前级
END_IF

(* —— 段 4：级数上限换算（级步换算，R28-2 两点向量） —— *)
IF NOT _bCfgBad THEN
    _nStageMax := TRUNC(fReheatMaxPct / fReheatStageStepPct);   // 级数上限（整除点精确取整，不越级）
    IF DINT_TO_REAL(DINT(_nStageMax)) * fReheatStageStepPct < fReheatMaxPct THEN
        _nStageMax := _nStageMax + 1;   // 余量进位到覆盖上限（上限 +1 向量：取整后余量补一级）
    END_IF
END_IF

(* —— 段 5：期望级数解算（温度需求 + 风量降档 + 互锁全关） —— *)
IF (NOT _bCfgBad) AND (NOT _bSigBad) THEN
    _rErr := fZoneSetC - fZoneTempC;                 // 温度偏差（> 0 需加热）
    IF bReheatInhibit THEN
        _nStageDes := 0;                             // 互锁：再热全关（规格强制）
        _uInfo := 16#0006_04B2;                      // 信息级：互锁生效
    ELSIF fAirflowPct < fMinAirflowPct THEN
        _nStageDes := 0;                             // 风量不足：按级降档目标（逐级走）
        _bLimitHold := TRUE;                         // 约束保持量
    ELSE
        IF _rErr > 0.5 THEN
            _nStageDes := _nStageMax;                // 明显需热：目标满级（级间延时节流逐级逼近）
        ELSIF _rErr < -0.5 THEN
            _nStageDes := 0;                         // 过热：目标 0 级
        ELSE
            _nStageDes := _nStage;                   // 死区内：维持当前级
        END_IF
    END_IF
END_IF

(* —— 段 6：级间延时节流推进（每 tStageDelay 向期望级走一级，防级联抖动） —— *)
IF (NOT _bCfgBad) AND (NOT _bSigBad) AND (_nStageDes <> _nStage) THEN
    IF tonStageDly.Q THEN
        _bStageBrk := TRUE;                          // 断输入请求：窗重开（自复位范式）
        IF _nStageDes > _nStage THEN
            _nStage := MIN(_nStage + 1, _nStageMax); // 升一级（上限钳制）
        ELSE
            _nStage := MAX(_nStage - 1, 0);          // 降一级（下界钳制）
        END_IF
    END_IF
END_IF

(* —— 段 7：出口单点映射（名实同源；每拍重算，无锁存码回放需求） —— *)
nActiveStage := _nStage;                             // 级数出口
fReheatCmdPct := DINT_TO_REAL(DINT(_nStage)) * fReheatStageStepPct;   // 再热输出 = 级数 × 级步
fReheatCmdPct := MIN(MAX(fReheatCmdPct, 0.0), fReheatMaxPct);         // 钳 [0, 上限]（禁越上界）
bMinAirflowLimit := _bLimitHold AND (fAirflowPct < fMinAirflowPct);   // 约束出口（每拍重算，解除式）
bReheatInhibitActive := bReheatInhibit AND (NOT _bCfgBad);            // 互锁镜像出口
IF _bCfgBad THEN
    nErrId := 16#0006_02B2;              // 故障级：组态非法（每拍重申）
    fReheatCmdPct := 0.0;                // 组态错输出全关（安全侧）
    nActiveStage := 0;
ELSIF bReheatInhibit THEN
    nErrId := 16#0006_04B2;              // 信息级：互锁全关
ELSIF _bSigBad THEN
    nErrId := 16#0006_01B2;              // 信息级：信号坏保持当前级
ELSIF bMinAirflowLimit THEN
    nErrId := 16#0006_03B2;              // 信息级：最小风量约束
END_IF

END_FUNCTION_BLOCK

(* ---- FB_DL_ThickenerFlocDoseCtrl.st ---- *)
(*
  Name: FB_DL_ThickenerFlocDoseCtrl
  Category: DL_Process
  Version: 1.0.0
  Round: R89 / 2026-11-25
  开源溯源：clean-room 自研（族 矿山破碎筛分，ST 开源生态实测 0 命中，无外部代码引入）
  功能：浓密机絮凝剂投加控制：给矿量前馈（g/t 基准投加）乘底流浓度反馈修正因子，输出溶液投加流量。
  边界条件：① 六入参全部过非有限闸；配置越域进冻结分支：输出保持上一有效值 + xValid = FALSE（R191 已声明）；
            ② xEnable = FALSE 语义：冻结保持末值（不降级为 0，避免投加泵被清零误动作），xValid 同拍置 FALSE；
            ③ 抗积分饱和：本件为乘性修正（无积分器，故无 windup 通路），修正因子钳位 0.7~1.4；
               输出达上限时冻结因子更新（保持末值），防止饱和期内因子持续堆高；
            ④ 固体吨位为代理量：以底流浓度近似给矿固体含量（保守偏小），代理假设见功能段。
  量纲自证：Q[m3/h] × ρ[t/m3] × C[−] = t/h；t/h × g/t = g/h；g/h ÷ g/L = L/h。
*)
FUNCTION_BLOCK FB_DL_ThickenerFlocDoseCtrl
VAR_INPUT
    xEnable : BOOL;             (* 投加使能 [-] Dosing enable *)
    fFeedM3h : REAL;            (* 给矿浆体流量 [m3/h] Feed slurry flow [m3/h] *)
    fDoseGpt : REAL;            (* 基准投加量（每吨固体） [g/t] Base dosage per tonne solids [g/t] *)
    fUnderDensityPct : REAL;    (* 底流浓度实测 [%] Underflow density actual [%] *)
    fUnderDensitySpPct : REAL;  (* 底流浓度设定 [%] Underflow density setpoint [%] *)
    fDoseMaxLph : REAL;         (* 投加泵流量上限 [L/h] Dosage pump ceiling [L/h] *)
END_VAR
VAR_OUTPUT
    fDoseLph : REAL;            (* 投加溶液流量 [L/h] Dosing solution flow [L/h] *)
    xSaturated : BOOL;          (* 输出已达上限 [-] Output saturated *)
    xValid : BOOL;              (* 配置与链路有效 [-] Configuration and chain valid *)
END_VAR
VAR
    _bInit : BOOL := FALSE;     (* 首扫初始化标志 [-] First-scan init flag *)
    _bCfgBad : BOOL := FALSE;   (* 配置非法当拍量 [-] Configuration bad *)
    _bCalcOk : BOOL := FALSE;   (* 本拍计算有效 [-] Calculation valid this scan *)
    _fTrim : REAL := 1.0;       (* 反馈修正因子（钳 0.7~1.4） [-] Feedback trim factor *)
    _fTrimNew : REAL := 1.0;    (* 本拍候选修正因子 [-] Candidate trim factor *)
    _fErrPct : REAL := 0.0;     (* 浓度偏差（设定 − 实测） [%] Density deviation [%] *)
    _fSolidsTph : REAL := 0.0;  (* 固体吨位代理量 [t/h] Solids tonnage proxy [t/h] *)
    _fDose : REAL := 0.0;       (* 投加流量保持量 [L/h] Dosing flow hold [L/h] *)
    _bSat : BOOL := FALSE;      (* 饱和锁存 [-] Saturation latch *)
END_VAR
VAR CONSTANT
    DL_EPS : REAL := 1.0E-9;        (* 除零判定容差 [-] Divide-by-zero tolerance *)
    DL_RHO_SL : REAL := 1.05;       (* 浆体密度代理值 [t/m3] Slurry density proxy [t/m3] *)
    DL_GPL : REAL := 0.5;           (* 絮凝剂溶液浓度 [g/L] Flocculant solution strength [g/L] *)
    DL_KFB : REAL := 0.5;           (* 反馈修正增益 [-] Feedback trim gain *)
    DL_TRIM_LO : REAL := 0.7;       (* 修正因子下限 [-] Trim floor *)
    DL_TRIM_HI : REAL := 1.4;       (* 修正因子上限 [-] Trim ceiling *)
    DL_PCT : REAL := 100.0;         (* 百分数基准 [%] Percent base *)
END_VAR
(* 首扫初始化：修正因子起点 1.0（纯前馈） *)
IF NOT _bInit THEN
    _fTrim := 1.0;
    _fDose := 0.0;
    _bSat := FALSE;
    _bInit := TRUE;
END_IF
(* 非有限闸（NaN 自反 + Inf 差值自减）+ 静态组态域闸：五浮点入参全枚举（R272） *)
_bCfgBad := (fFeedM3h <> fFeedM3h) OR ((fFeedM3h - fFeedM3h) <> 0.0)
         OR (fDoseGpt <> fDoseGpt) OR ((fDoseGpt - fDoseGpt) <> 0.0)
         OR (fUnderDensityPct <> fUnderDensityPct) OR ((fUnderDensityPct - fUnderDensityPct) <> 0.0)
         OR (fUnderDensitySpPct <> fUnderDensitySpPct) OR ((fUnderDensitySpPct - fUnderDensitySpPct) <> 0.0)
         OR (fDoseMaxLph <> fDoseMaxLph) OR ((fDoseMaxLph - fDoseMaxLph) <> 0.0)
         OR (fFeedM3h < 0.0) OR (fFeedM3h > 5000.0)
         OR (fDoseGpt < 1.0) OR (fDoseGpt > 500.0)
         OR (fUnderDensityPct < 0.0) OR (fUnderDensityPct > 60.0)
         OR (fUnderDensitySpPct < 5.0) OR (fUnderDensitySpPct > 60.0)
         OR (fDoseMaxLph < 0.1) OR (fDoseMaxLph > 5000.0);
_bCalcOk := xEnable AND (NOT _bCfgBad);
IF _bCalcOk THEN
    (* 固体吨位代理：Q[m3/h] × ρ[t/m3] × C[−] = t/h *)
    _fSolidsTph := fFeedM3h * DL_RHO_SL * (fUnderDensityPct / DL_PCT);
    (* 偏差：设定 − 实测，正值表示底流偏稀需加大投加 *)
    _fErrPct := fUnderDensitySpPct - fUnderDensityPct;
    (* 候选修正因子 + 钳位（量值饱和；饱和期间冻结更新以抗饱和） *)
    IF NOT _bSat THEN
        _fTrimNew := 1.0 + DL_KFB * (_fErrPct / DL_PCT);
        IF _fTrimNew < DL_TRIM_LO THEN
            _fTrimNew := DL_TRIM_LO;
        ELSIF _fTrimNew > DL_TRIM_HI THEN
            _fTrimNew := DL_TRIM_HI;
        END_IF
        _fTrim := _fTrimNew;
    END_IF
    (* 前馈 × 反馈：t/h × g/t = g/h；÷ g/L = L/h *)
    _fDose := ((_fSolidsTph * fDoseGpt) * _fTrim) / DL_GPL;
    (* 上限钳位：达上限即置饱和并冻结因子，防饱和期堆高 *)
    IF _fDose >= fDoseMaxLph THEN
        _fDose := fDoseMaxLph;
        _bSat := TRUE;
    ELSE
        _bSat := FALSE;
    END_IF
END_IF
(* 统一出口（单点赋值）：冻结分支保持上一有效值，保持量来源均为已过闸的有限值（R273） *)
fDoseLph := _fDose;
xSaturated := _bSat AND _bCalcOk;
xValid := _bCalcOk;
END_FUNCTION_BLOCK
